// TwinCAT 3 PLC project axis_4
// ProgramVersion: 3.1.4026.27
// libraries:
//   Tc2_MC2, * (Beckhoff Automation GmbH)
//   Tc2_Standard, * (Beckhoff Automation GmbH)
//   Tc2_System, * (Beckhoff Automation GmbH)
// project tree:
//   DUTs/ ST_AxisMonitor.TcDUT, ST_MachineMonitor.TcDUT, ST_AxisCommand.TcDUT, ST_ControlStation.TcDUT, ST_AxisConfig.TcDUT, ST_TrajectoryPoint.TcDUT, ST_AxisAds.TcDUT
//   GVLs/ GVL_control.TcGVL, GVL_HMI.TcGVL, GVL_motion.TcGVL, GVL_sy.TcGVL, GVL_axis.TcGVL
//   POUs/ControlAuthority_控制权/ F_ControlDecision.TcPOU, FB_ControlAuthority.TcPOU
//   POUs/ManualControl_手动控制/ FB_AxisCommandGate.TcPOU, FB_AxisControl.TcPOU
//   POUs/Feedback_反馈/ FB_HmiFeedback.TcPOU
//   POUs/AxisConfig_轴配置/ F_AxisPositionValid.TcPOU, F_AxisConfigValid.TcPOU, FB_AxisConfig.TcPOU
//   POUs/Trajectory_点位与轨迹/ FB_FourAxisTrajectory.TcPOU, F_TrajectoryPoint.TcPOU
//   / PlcTask.TcTTO
//   POUs/ MAIN.TcPOU
// real-time tasks:
//   TASK PlcTask: cycle T#10ms, priority 20, ADS port 350
//   TASK PlcTask1: cycle T#2ms, priority 7, ADS port 351
// motion (NC):
//   TASK NC-Task 1 SAF: cycle T#2ms, priority 4, ADS port 501
//   TASK NC-Task 1 SVB: cycle T#10ms, priority 8, ADS port 511
//   AXIS axis1 (id 1)
//     OtherSettings: AllowMotionCmdToSlave=true
//     encoder EncType=19
//       EncPara: MaxCount=#xffffffff
//     drive DrvType=16
//       DrvPara: MaxCount=#xffffffff
//         Analog: TorqueSetpointScale=10, ScaleFactorActTorque=0.1
//         TimeComp: TaskDelayCycles=1
//     controller CtrType=1
//       CtrPara: PriorControlFactor=1
//         Observer: BandWidth=20
//   AXIS axis2 (id 2)
//     OtherSettings: AllowMotionCmdToSlave=true
//     encoder EncType=19
//       EncPara: MaxCount=#xffffffff
//     drive DrvType=16
//       DrvPara: MaxCount=#xffffffff
//         Analog: TorqueSetpointScale=10, ScaleFactorActTorque=0.1
//         TimeComp: TaskDelayCycles=1
//     controller CtrType=1
//       CtrPara: PriorControlFactor=1
//         Observer: BandWidth=20
//   AXIS axis3 (id 3)
//     OtherSettings: AllowMotionCmdToSlave=true
//     encoder EncType=19
//       EncPara: MaxCount=#xffffffff
//     drive DrvType=16
//       DrvPara: MaxCount=#xffffffff
//         Analog: TorqueSetpointScale=10, ScaleFactorActTorque=0.1
//         TimeComp: TaskDelayCycles=1
//     controller CtrType=1
//       CtrPara: PriorControlFactor=1
//         Observer: BandWidth=20
//   AXIS axis4 (id 4)
//     OtherSettings: AllowMotionCmdToSlave=true
//     encoder EncType=19
//       EncPara: MaxCount=#xffffffff
//     drive DrvType=16
//       DrvPara: MaxCount=#xffffffff
//         Analog: TorqueSetpointScale=10, ScaleFactorActTorque=0.1
//         TimeComp: TaskDelayCycles=1
//     controller CtrType=1
//       CtrPara: PriorControlFactor=1
//         Observer: BandWidth=20
// variable links:
//   axis_4/axis_4 Instance <-> NC-Task 1 SAF/Axes/axis1
//     PlcTask Inputs/GVL_sy.axis[1].NcToPlc <-> 输出/ToPlc
//     PlcTask Outputs/GVL_sy.axis[1].PlcToNc <-> 输入/FromPlc
//   axis_4/axis_4 Instance <-> NC-Task 1 SAF/Axes/axis2
//     PlcTask Inputs/GVL_sy.axis[2].NcToPlc <-> 输出/ToPlc
//     PlcTask Outputs/GVL_sy.axis[2].PlcToNc <-> 输入/FromPlc
//   axis_4/axis_4 Instance <-> NC-Task 1 SAF/Axes/axis3
//     PlcTask Inputs/GVL_sy.axis[3].NcToPlc <-> 输出/ToPlc
//     PlcTask Outputs/GVL_sy.axis[3].PlcToNc <-> 输入/FromPlc
//   axis_4/axis_4 Instance <-> NC-Task 1 SAF/Axes/axis4
//     PlcTask Inputs/GVL_sy.axis[4].NcToPlc <-> 输出/ToPlc
//     PlcTask Outputs/GVL_sy.axis[4].PlcToNc <-> 输入/FromPlc

CONFIGURATION axis_4
    RESOURCE PLC ON TwinCAT3
        TASK PlcTask(INTERVAL := T#2ms, PRIORITY := 7);
        PROGRAM MAIN WITH PlcTask : MAIN;
    END_RESOURCE
END_CONFIGURATION

// ---- DUTs/ST_AxisMonitor.TcDUT
{attribute 'pack_mode' := '1'}
TYPE ST_AxisMonitor :
STRUCT
    // 仅反馈，固定 22 字节；顺序与 C# PlcAxisMonitor 完全一致。
    lrActualPosition : LREAL; // PLC 从基础轴转发、上位机只读：NC 实际位置，单位跟随 NC，现场单位尚未确认。
    lrSpeed : LREAL; // PLC 从基础轴转发、上位机只读：NC 实际速度，单位为 NC 位置单位/秒，含方向正负号。
    xHomed : BOOL; // PLC 从基础轴转发、上位机只读：NC 已回原反馈，不是回原请求。
    xError : BOOL; // PLC 从基础轴转发、上位机只读：本轴 NC 或基础 MC 功能块错误。
    xPositiveLimit : BOOL; // PLC 从基础轴转发、上位机只读：正向硬限位或 NC 正向软限位超限。
    xNegativeLimit : BOOL; // PLC 从基础轴转发、上位机只读：负向硬限位或 NC 负向软限位超限。
    xOriginSignal : BOOL; // PLC 从基础轴转发、上位机只读：原点传感器信号，不代表回原已经完成。
    xEnabled : BOOL; // MC_Power.Status，使能反馈，不以运动位代替。 PLC 从基础轴转发，上位机只读。
END_STRUCT
END_TYPE

// ---- DUTs/ST_MachineMonitor.TcDUT
{attribute 'pack_mode' := '1'}
TYPE ST_MachineMonitor :
STRUCT
    // 布局版本 4，总长 164 字节；修改字段时须同步上位机并升级版本。
    nVersion : UINT; // PLC 写、上位机只读：监控协议布局版本，当前为 4，上位机据此校验帧。
    nByteSize : UINT; // PLC 写、上位机只读：完整监控结构字节数，当前为 164，不是轴数量或有效点数。
    nControlOwner : UINT; // PLC 写、上位机只读：仲裁持有者，0 未分配、1 造波控制室、2 拖车本地、3 远程操作室。
    nControlMode : UINT; // PLC 写、上位机只读：0 未分配、1 手动、2 轨迹占用；由持有者和轨迹 Busy 推导，不是模式请求。
    nWaveState : UINT; // PLC 写、上位机只读：页面状态 0 待机、1 准备、2 运行、4 停止中、5 已停止、6 完成、7 故障。
    uiWaveFaultCode : UINT; // PLC 写、上位机只读：组或首个轴的 16 位显示错误码，超过 65535 显示 65535；完整码见 GVL_HMI.udiDetailedFaultCode。
    udiHeartbeat : UDINT; // PLC 每约 500 ms 递增的反馈心跳，溢出回 0；上位机据变化判断反馈新鲜度，不由上位机写。
    Axis1 : ST_AxisMonitor; // PLC 写、上位机只读：NC 轴 1 的实际反馈，布局固定为 ST_AxisMonitor。
    Axis2 : ST_AxisMonitor; // PLC 写、上位机只读：NC 轴 2 的实际反馈，布局固定为 ST_AxisMonitor。
    Axis3 : ST_AxisMonitor; // PLC 写、上位机只读：NC 轴 3 的实际反馈，布局固定为 ST_AxisMonitor。
    Axis4 : ST_AxisMonitor; // PLC 写、上位机只读：NC 轴 4 的实际反馈，布局固定为 ST_AxisMonitor。
    // 轨迹及自动准备反馈，顺序对应 C#，继续 1 字节对齐。
    nTrajectoryState : UINT; // PLC 写、上位机只读：轨迹内部状态 0空闲/5拼表/10校验/15首点定位/20开外部给定/30运行/40末点保持/50减速/60关给定/70等停稳/90故障。
    nReceivedCount : UDINT; // PLC 写、上位机只读：四轴已登记接收的点数，也是下段起始偏移；不是已拼表点数。
    nLoadedCount : UDINT; // PLC 写、上位机只读：四轴均已拼入执行表的点数；不代表已校验通过或已运动完成。
    nPointCount : UDINT; // PLC 转发、上位机只读：上位机在 GVL_motion 中声明的目标总点数，不等于已接收或已拼接点数。
    nCurrentPoint : UDINT; // PLC 写、上位机只读：最近准备送给 NC 的点号，从 0 开始；不表示实际轴已到该点。
    udiReceivedSequence : UDINT; // PLC 写、上位机只读：当前接收表所属轨迹序号，清表后为 0；用于核对收段确认。
    udiAcceptedSequence : UDINT; // PLC 写、上位机只读：已校验通过并进入首点定位的轨迹序号，用于防止重复执行，不是完成序号。
    udiErrorId : UDINT; // PLC 写、上位机只读：轨迹块完整诊断码或 MC 原始 ErrorID；不汇总单轴错误，0 表示当前无组错误码。
    nUploadStation : UINT; // PLC 写、上位机只读：接收表归属站，0 无归属、1..3 对应控制站；不是上位机直接申请的授权。
    xUploadBusy : BOOL; // PLC 写、上位机只读：状态 5 正在统一拼表；不表示上位机当前正在写 ADS。
    xDataReady : BOOL; // PLC 写、上位机只读：完整位置表已拼接就绪；数值由上位机预检，不代表轴已使能或已到首点。
    xTrajectoryBusy : BOOL; // PLC 写、上位机只读：状态 10..70 占用轴控制，包含启动检查、定位、运行和退出；拼表状态 5 不占用。
    xRunning : BOOL; // PLC 写、上位机只读：仅内部状态 30 正常取点运行，首点定位和减速退出不算正常取点。
    xDone : BOOL; // PLC 写、上位机只读：轨迹自然完成且退出后保持，不以启动写入成功或末点已发送代替。
    xError : BOOL; // PLC 写、上位机只读：轨迹组故障保持位，确认退出并满足静止条件后由组复位请求清除。
    xStopped : BOOL; // PLC 写、上位机只读：人工组停止流程完成后保持，区别于自然完成 xDone 和组故障 xError。
    xMotionPermit : BOOL; // PLC 写、上位机只读：当前运行许可反馈，不等于已获控制权、轴已使能或硬件安全确认。
    xConfigValid : BOOL; // PLC 写、上位机只读：四轴设备参数的监控校验结果；不表示已使能或轨迹整表已校验。
    xAxesIdle : BOOL; // PLC 写、上位机只读：四轴有效停稳、基础块空闲且无外部给定；未使能轴也可满足空闲。
    xAxisFault : BOOL; // PLC 写、上位机只读：任一基础轴错误、NC 错误或 NC I/O 无效；不是仅指驱动器报警。
    xAxesStopped : BOOL; // 实际停车完成；MC_Stop 可以尚未释放。 PLC 汇总四轴 xStopped，上位机只读；反馈无效时不能确认停稳。
    // 配套版本及首次故障；均由 PLC 写，上位机只读。
    udiProgramVersion : UDINT; // PLC 源码发布号，2026102301；下载后才更新在线值。
    nBehaviorVersion : UINT; // 1=上位机整表预检，PLC 保留接收协议与运动联锁。
    nFaultAxis : UINT; // 首次轨迹故障轴号 1..4，0 表示组条件或未定位到单轴。
    nFaultSource : UINT; // 首次故障来源，含联停条件和 MC 块，见故障说明。
    nFaultState : UINT; // 首次故障发生时的轨迹阶段，不随停车阶段变化。
    udiCleanupErrorId : UDINT; // 停车/关闭/退出的首个错误，不能覆盖原始轨迹故障。
END_STRUCT
END_TYPE

// ---- DUTs/ST_AxisCommand.TcDUT
TYPE ST_AxisCommand :
STRUCT
    // 单个站点的命令邮箱，不含反馈；本站上位机写请求，PLC 在控制权交接时清空旧命令。
    xStart : BOOL; // 本站上位机写：保持型使能请求，TRUE 请求使能、FALSE 请求撤使能；不是轨迹启动或实际使能反馈。
    xStop : BOOL; // 本站上位机写：保持型停止请求，TRUE 停车、FALSE 撤请求；当前客户端发送 50 ms 脉冲，停稳另读反馈。
    jogz : BOOL; // 本站上位机写：正向点动保持位，按下 TRUE、松开 FALSE；不是实际正转反馈。
    jogf : BOOL; // 本站上位机写：负向点动保持位，按下 TRUE、松开 FALSE；不是实际反转反馈。
    gohome : BOOL; // 本站上位机写：回原上升沿请求，须先回 FALSE 再次置 TRUE；当前客户端脉冲 50 ms。
    reset : BOOL; // 本站上位机写：轴故障复位上升沿请求，须先回 FALSE 再次置 TRUE；当前客户端脉冲 50 ms。
    lrJogSpeed : LREAL; // 本站上位机写：点动速度幅值，单位为 NC 位置单位/秒；启动点动前先写速度，再写方向位。
END_STRUCT
END_TYPE

// ---- DUTs/ST_ControlStation.TcDUT
TYPE ST_ControlStation :
STRUCT
    // 站点写：先写 nAction，再提交新的非零序号；心跳独立持续更新。
    udiHeartbeat : UDINT; // 本站上位机持续写变化计数，不是请求沿；PLC 见过变化后判在线，连续 3 秒不变判离线。
    nAction : UINT; // 1 申请，2 释放。 本站上位机先写动作，再更新请求序号；动作值本身不代表已获授权。
    udiRequestSequence : UDINT; // 本站上位机写：新的非零序号提交一次请求，PLC 按与应答序号不同识别新请求，不按 BOOL 上升沿。
    xWaveSession : BOOL; // 本站发送/自动准备/执行会话，锁住交接；失联后不再保留锁。 本站写保持位，PLC 在交接时清零；表示软件会话占用，不是实际轨迹运行反馈。
    aAxis : ARRAY[1..4] OF ST_AxisCommand; // 本站上位机写：固定对应轴 1..4 的手动命令；PLC 仅转交授权站，交接时清除各站旧命令。
    // PLC 写，站点只读：请求是否成功必须看同序号应答，不能以写成功代替授权。
    udiAckSequence : UDINT; // PLC 写、本站只读：已处理的请求序号，必须等于本次请求序号后才能采用 nResult。
    nResult : UINT; // 1 成功；2 运行锁定；3 保留（旧版现场授权拒绝）；4 离线；5 非持有者；6 优先级；7 无效操作。 PLC 写、本站只读；须结合本次相同序号的 udiAckSequence 判断。
    xOnline : BOOL; // PLC 写、本站只读：心跳变化及 3 秒超时判断结果；ADS 连接成功不等于本站在线。
    xGranted : BOOL; // PLC 写、本站只读：当前持有者且在线、未失联退出时为 TRUE；写请求成功不代表获授权。
END_STRUCT
END_TYPE

// ---- DUTs/ST_AxisConfig.TcDUT
TYPE ST_AxisConfig :
STRUCT
    // 单位跟随 NC：位置、位置/秒、位置/秒²。必须按设备行程填写。
    // 参数在 FB_AxisConfig 中集中填写到 GVL_motion.aConfig；当前值仅用于虚拟轴调试，现场位置单位尚未确认。
    lrMinPosition : LREAL; // 设备配置值，PLC 读取：最小允许位置边界，单位跟随 NC 位置单位。
    lrMaxPosition : LREAL; // 设备配置值，PLC 读取：最大允许位置边界，单位跟随 NC 位置单位，须大于最小位置。
    lrMaxVelocity : LREAL; // 设备配置值，PLC 读取：点动及轨迹的速度上限，正值，单位为 NC 位置单位/秒。
    lrMaxAcceleration : LREAL; // 设备配置值，PLC 读取：点动/定位加速度及轨迹加速度幅值上限，正值，单位为 NC 位置单位/秒²。
    lrStopDeceleration : LREAL; // 设备配置值，PLC 读取：手动、首点定位及轨迹停车减速度幅值，正值且不大于最大加速度，单位为 NC 位置单位/秒²。
    lrStartTolerance : LREAL; // 设备配置值，PLC 读取：首点定位完成后实际位置和设定位置到首点的容差，轨迹要求大于 0，单位跟随 NC。
    lrInitVelocity : LREAL; // 轨迹启动前，四轴各自移动到首点的速度。 配置方填写、PLC 读取；须大于 0 且不超过最大速度，单位为 NC 位置单位/秒。
END_STRUCT
END_TYPE

// ---- DUTs/ST_TrajectoryPoint.TcDUT
TYPE ST_TrajectoryPoint :
STRUCT
    // PLC 内部送点使用；上位机只下发 LREAL 位置表，速度/加速度由相邻点计算。
    lrPosition : LREAL; // PLC 内部绝对位置给定，来自当前表点或停车积分；不是实际位置反馈，单位跟随 NC。
    lrVelocity : LREAL; // PLC 内部速度给定，正常运行由相邻点按 2 ms 中心差分计算，首尾为 0；单位为 NC 位置单位/秒。
    lrAcceleration : LREAL; // PLC 内部加速度给定，正常运行由相邻点按 2 ms 二阶差分计算，停车时另算；单位为 NC 位置单位/秒²。
END_STRUCT
END_TYPE

// ---- DUTs/ST_AxisAds.TcDUT
TYPE ST_AxisAds :
STRUCT
    // PLC → 上位机：反馈量
    lrActualPosition : LREAL; // PLC 写、上位机只读：NC 实际位置，单位跟随 NC 位置单位，现场尚未确认。
    lrSpeed          : LREAL; // PLC 写、上位机只读：NC 实际速度，单位为 NC 位置单位/秒，正负号表示方向。
    xMotorRun        : BOOL; // PLC 写、上位机只读：NC Moving 实际运动位，不是使能成功或运动请求。
    xHomed           : BOOL; // PLC 写、上位机只读：NC Homed 回原有效反馈，不以 gohome 请求代替。
    xError           : BOOL; // PLC 写、上位机只读：NC 或 Power/Stop/Home/Jog/Reset 任一错误，错误码见 udiErrorId。
    xPositiveLimit   : BOOL; // PLC 写、上位机只读：正向硬限位或 NC 正向软限位超限，TRUE 表示触发。
    xNegativeLimit   : BOOL; // PLC 写、上位机只读：负向硬限位或 NC 负向软限位超限，TRUE 表示触发。
    xOriginSignal    : BOOL; // PLC 写、上位机只读：实际原点传感器信号，不等于已完成回原。

    // PLC 命令门转交授权站的命令；上位机应写 aStation[本站].aAxis，不直写以下字段。
    xStart     : BOOL; // PLC 命令门转交：保持型使能请求，TRUE 请求使能、FALSE 先停车再撤使能；实际结果看 xEnabled。
    xStop      : BOOL; // PLC 命令门转交：保持型停止请求，TRUE 请求停车并维持停止条件，FALSE 撤请求；完成看 xStopped。
    jogz       : BOOL; // PLC 命令门转交：正向点动保持请求，按下 TRUE、释放 FALSE 后减速；与 jogf 同时 TRUE 不点动。
    jogf       : BOOL; // PLC 命令门转交：负向点动保持请求，按下 TRUE、释放 FALSE 后减速；与 jogz 同时 TRUE 不点动。
    gohome     : BOOL; // PLC 命令门转交：回原上升沿请求，须回 FALSE 后才能再次触发；完成看 xHomed。
    reset      : BOOL; // PLC 命令门转交：轴故障复位上升沿请求，须回 FALSE 后再次触发；故障是否消除看 xError。
    lrJogSpeed : LREAL; // PLC 命令门转交：点动速度幅值，单位为 NC 位置单位/秒，须大于 0 且不超过配置上限。
    // 新字段放在末尾；上位机应按 ADS 符号访问，整结构读写须同步更新布局。
    xEnabled : BOOL; // MC_Power.Status，使能反馈；xStart 为保持型使能请求。 PLC 每扫描写，上位机只读。
    xBusy : BOOL; // PLC 写、上位机只读：轨迹占用或 Jog/Home/Stop/Reset 忙，含停止锁保持，不等于轴正在运动。
    xStopped : BOOL; // 实际停稳且回原/点动退出，允许 MC_Stop.Done 保持。 PLC 写、上位机只读；不是停止请求，也不要求停止锁已经释放。
    udiErrorId : UDINT; // PLC 写、上位机只读：按 NC/Power/Stop/Home/Jog/Reset 顺序取首个错误码，0 表示未发布错误码。
END_STRUCT
END_TYPE

// ---- GVLs/GVL_control.TcGVL
{attribute 'qualified_only'}
VAR_GLOBAL
    // 新三站协议编码：1 造波控制室，2 拖车本地，3 远程操作室；数字小优先级高。
    // 各站只写自己的请求、心跳和手动命令；应答与授权结果由 PLC 写。
    aStation : ARRAY[1..3] OF ST_ControlStation; // 三站独立邮箱；各站写自己的请求/心跳/命令，PLC 写应答与授权反馈。
    // 纯软件申请，不使用现场主控选择位；PLC 按心跳、运行锁及优先级授予控制权。
    // 以下由仲裁块写，任何上位机都不能直接写 Owner 来取得权限。
    nOwner : UINT; // PLC 发布的持有站：0 未分配，1 控制室、2 拖车本地、3 远程室；上位机只读。
    xLocked : BOOL; // 统一交接锁：运动、待执行运动命令，或 I/O 故障下轴仍使能。
    xCanRelease : BOOL; // 由 Owner 和 xLocked 推导，保留此反馈供已有上位机兼容。
    xFeedbackInvalid : BOOL; // 任一轴 NC I/O 无效；单独提示，基础轴块禁止新使能/运动。
    xCanCommand : BOOL; // PLC 发布的当前持有站命令许可；需持有站在线且未失联锁存。
    xOwnerChanged : BOOL; // 本扫描发生交接或撤权重授的标志，用于清旧命令、阻止同扫描重放。
    xStopOwner : BOOL; // 失联后撤销命令并停车，保持旧 Owner 直到停稳。
END_VAR

// ---- GVLs/GVL_HMI.TcGVL
{attribute 'qualified_only'}
VAR_GLOBAL
    // 整块只读监控接口；由 FB_HmiFeedback 在轴块执行后发布。
    stMonitor : ST_MachineMonitor; // PLC 每扫描发布的整块只读监控帧，包含四轴实际状态与组反馈。
    // 保留完整故障码及轨迹诊断；全部由 PLC 发布，上位机只读。
    udiDetailedFaultCode : UDINT; // 完整错误码，不丢失高 16 位。
    nFaultAxis : UINT; // 0 为组故障或无错误；1..4 为对应轴的首个错误。
    nTrajectoryState : UINT; // 轨迹块内部 nState，区别于上述页面状态编码。
    nCurrentPoint : UDINT; // PLC 发布的最近外部给定点号，从 0 开始，不表示机械轴实际到位。
    nLoadedCount : UDINT; // PLC 发布的四轴已拼入执行表的点数。
    nPointCount : UDINT; // PLC 发布的目标单轴总点数，不表示接收或执行进度。
    xDataReady : BOOL; // PLC 发布的整表拼接完成标志，不表示数值校验或首点定位完成。
    xTrajectoryBusy : BOOL; // PLC 发布的轨迹占轴标志，含校验、定位、执行和退出阶段。
END_VAR

// ---- GVLs/GVL_motion.TcGVL
{attribute 'qualified_only'}
// ADS 协议：上位机写命令/数据，PLC 写反馈；状态字段只供上位机读取。
// PC 连续提交各段，全部下发后用 xAssemble 请求 PLC 拼表；xDataReady 后才允许启动。
// xUpload/xAssemble/xClear/xStart/xReset 都需回 FALSE 后再产生下一次上升沿。
VAR_GLOBAL
    // 运行许可由 MAIN 每扫描写入；当前仅用于虚拟轴调试。
    xMotionPermit : BOOL; // 实机改接安全继电器允许反馈，不代替硬件安全回路。
    axPositiveLimit : ARRAY[1..4] OF BOOL; // 四轴正向硬限位输入，索引为轴号 1～4，TRUE 表示触发。
    axNegativeLimit : ARRAY[1..4] OF BOOL; // 四轴负向硬限位输入，索引为轴号 1～4，TRUE 表示触发。
    axHomeSensor : ARRAY[1..4] OF BOOL; // 四轴原点开关输入，索引为轴号 1～4，传给 NC 标准回零校准凸轮。
    // 四轴配置只在 FB_AxisConfig 中填写，手动、反馈和轨迹均读取此数组。
    aConfig : ARRAY[1..4] OF ST_AxisConfig; // 单位跟随 NC；空闲时由配置块直接更新，运动期间保持。

    // 以下为上位机写入的轨迹命令与点位；nUploadStation、xStopped 两项由 PLC 写、上位机只读。
    nCommandStation : UINT; // 上位机命令来源，必须等于有效 Owner；不是授权本身。
    nUploadStation : UINT; // PLC 锁存的上传所属站，只读。
    xStopped : BOOL; // 人工停止完成；不同于自然完成 xDone 或故障。
    // 参考旧工程的独立分段区：21 段、每段四轴、每轴最多 100000 个 LREAL 点。
    // 下标依次为 [段号, 轴号, 段内点号]；已提交段禁止覆盖，全部下发后统一拼接。
    aUpload : ARRAY[0..20, 1..4, 0..99999] OF LREAL; // 上位机写入的独立位置段：[段0～20,轴1～4,段内点0～99999]，数值单位跟随 NC。
    nPointCount : UDINT; // 整条轨迹总点数，4..2100000。
    nSampleTimeUs : UINT := 2000; // 单位微秒，目前仅接受 2000。
    udiUploadSequence : UDINT; // 整条轨迹使用同一个非零序号。
    nUploadOffset : UDINT; // 本段全局偏移，必须等于 nReceivedCount，段号=偏移/100000。
    nUploadCount : UDINT; // 非末段必须 100000 点；末段为总点数的剩余量。
    xUpload : BOOL; // 四轴本段数据写完后上升沿登记，只确认接收，不拼表。
    xAssemble : BOOL; // 全部段确认后上升沿请求统一拼表；拼接期间所有段保持不变。
    xClear : BOOL; // 空闲时上升沿清除整条位置表的就绪状态，开始新一轮上传。
    xStart : BOOL; // 完整位置表到齐后，上升沿启动。
    xStop : BOOL; // 保持型组停止，启动前必须释放。
    xReset : BOOL; // 清组故障；各轴故障用 Axis1..4.reset。
    udiHeartbeat : UDINT; // 校验/运动期间 1 秒不变化则联停。

    // 以下字段由 PLC 写，上位机只读。
    nReceivedCount : UDINT; // 已登记的下发点数，也是下一段允许的起始偏移；不代表已拼接。
    udiReceivedSequence : UDINT; // 已登记各段所属轨迹序号，清表后为 0。
    xUploadBusy : BOOL; // 全部下发后的统一拼表正在执行，不表示 PC 正在写 ADS。
    nLoadedCount : UDINT; // 四轴均已拼入完整表的点数；下发期间始终为 0。
    xDataReady : BOOL; // 全部段已统一拼接完成，不表示已校验或已定位到首点。
    xBusy : BOOL; // 校验、首点定位、执行和退出期间占用轴控制。
    xRunning : BOOL; // 状态 30，首点定位及减速不算正常取点运行。
    xDone : BOOL; // 正常完成后保持，清表/复位/新启动时清除。
    xError : BOOL; // 组故障保持位，需确认退出和静止后复位。
    udiErrorId : UDINT; // 首次故障的程序诊断码或 MC 原始 ErrorID，详见说明文档。
    nFaultAxis : UINT; // 首次故障轴 1..4；组故障或无故障为 0，复位时清除。
    nFaultSource : UINT; // 首次故障来源：1许可/2控制权/3使能/4单轴停止/5手动冲突/6限位，7..20见故障说明。
    nFaultState : UINT; // 首次故障发生阶段；故障退出期间保持，不能用当前停车阶段替代。
    udiCleanupErrorId : UDINT; // 首个停车、关闭或退出错误，保留原始 udiErrorId。
    nState : UINT; // 对应轨迹块 CASE 的 0/5/10/15/20/30/40/50/60/70/90。
    nCurrentPoint : UDINT; // 最近送出的点号，0 起始。
    udiAcceptedSequence : UDINT; // 已进入首点定位的轨迹序号，不能重复执行。
END_VAR

// ---- GVLs/GVL_sy.TcGVL
VAR_GLOBAL

axis  : ARRAY[1..4] OF AXIS_REF; // 四根 NC 轴引用，固定索引 1～4；轴状态从 NC 读取，运动块经此接口下发控制。

END_VAR

// ---- GVLs/GVL_axis.TcGVL
VAR_GLOBAL
    // PLC 内部手动命令与轴反馈；命令由 A03_ManualCommands 转交，反馈由基础轴块更新。
    // 上位机手动命令写 GVL_control.aStation[站号].aAxis，状态读取 GVL_HMI.stMonitor。

    Axis1 : ST_AxisAds; // 轴1内部手动命令与实际反馈；命令由命令门转交，反馈由轴1基础块更新。
    Axis2 : ST_AxisAds; // 轴2内部手动命令与实际反馈；命令由命令门转交，反馈由轴2基础块更新。
    Axis3 : ST_AxisAds; // 轴3内部手动命令与实际反馈；命令由命令门转交，反馈由轴3基础块更新。
    Axis4 : ST_AxisAds; // 轴4内部手动命令与实际反馈；命令由命令门转交，反馈由轴4基础块更新。


END_VAR

// ---- POUs/MAIN.TcPOU
// PlcTask 每 2 ms 调用；先刷新反馈，再判组条件，再轨迹，最后基础轴块。
// 每轴的 NC 引用、ADS 数据、参数及传感器索引必须一一对应。
PROGRAM MAIN
VAR
    fbAxisConfig : FB_AxisConfig; // 独立轴配置入口，仅在有效空闲时应用本块的虚拟轴参数。
    fbAxis1 : FB_AxisControl; // 轴1基础控制实例，固定对应 GVL_sy.axis[1] 和 GVL_axis.Axis1。
    fbAxis2 : FB_AxisControl; // 轴2基础控制实例，固定对应 GVL_sy.axis[2] 和 GVL_axis.Axis2。
    fbAxis3 : FB_AxisControl; // 轴3基础控制实例，固定对应 GVL_sy.axis[3] 和 GVL_axis.Axis3。
    fbAxis4 : FB_AxisControl; // 轴4基础控制实例，固定对应 GVL_sy.axis[4] 和 GVL_axis.Axis4。
    fbAuthority : FB_ControlAuthority; // 三站控制权仲裁实例，处理申请、释放、心跳和交接锁。
    aCommandGate : ARRAY[1..4] OF FB_AxisCommandGate; // 四轴手动命令门，只向对应轴转交当前持有站的有效命令。
    xControlBusy : BOOL; // 实际运动、轨迹或轴块忙的汇总，作为禁止控制权交接的判据。
    nManualStation : UINT; // 本扫描允许读取的站号；0 时命令门清除旧请求。
    fbTrajectory : FB_FourAxisTrajectory; // 四轴点位接收、拼表、校验及轨迹执行实例。
    fbHmiFeedback : FB_HmiFeedback; // 四轴执行结果发布到 switch 只读监控接口。
    xAllEnabled : BOOL; // 四轴使能反馈，用于运行中判断是否掉使能。
    xAxesReady : BOOL; // 轨迹启动就绪：四轴使能、回原、静止且不在停车。
    nAbortReason : UINT; // 本扫描首个联停原因；0 表示没有联停请求。
    xAbort : BOOL; // 整组联停请求，汇总许可丢失、撤使能、命令冲突及限位等条件。
    xAxisFault : BOOL; // 任一基础轴错误或 NC 错误、I/O 无效，供轨迹块判断故障。
    i : INT; // 四轴状态汇总的循环轴号，范围 1～4。
END_VAR

// 当前仅用于虚拟轴软件调试，明确给出运行许可。
// 接实机前必须将下一行替换为现场安全继电器的运行允许反馈。
GVL_motion.xMotionPermit := TRUE;

// 刷新四轴实际状态；只读取 NC 反馈，不要求持有控制权。
A01_ReadAxisStatus();

// 汇总交接条件并处理控制权；写入 GVL_control 仲裁反馈。
A02_ControlAuthority();

// 轴配置单独处理，使用当前运动锁和现有空闲反馈。
fbAxisConfig();

// 取出授权站手动命令；通过命令门写入 GVL_axis 命令字段。
A03_ManualCommands();

// 汇总轨迹联锁并调用原轨迹块；更新 GVL_motion 轨迹状态。
A04_TrajectoryControl();

// 调用四轴基础控制；更新 NC 控制输出及 GVL_axis 实际反馈。
A05_ManualAxes();

// 发布本扫描执行后的反馈；只写 GVL_HMI，不产生运动命令。
A06_PublishFeedback();

ACTION A01_ReadAxisStatus:
// 刷新四轴实际状态；只读取 NC 反馈，不要求持有控制权。
// 先统一刷新轴状态，再决定四轴本周期的共同轨迹帧。
FOR i := 1 TO 4 DO
 GVL_sy.axis[i].ReadStatus();
 END_FOR
END_ACTION

ACTION A02_ControlAuthority:
// 汇总交接条件并处理控制权；写入 GVL_control 仲裁反馈。
// 运行锁：点动、回原、轨迹、停止/退出及未消费的运动命令都阻止交接。
// 使用 NC 状态、实际速度和轴块 Busy；I/O 无效单独发布，不能冒充运动占用。
xControlBusy := GVL_motion.xBusy OR GVL_axis.Axis1.xBusy OR GVL_axis.Axis2.xBusy
    OR GVL_axis.Axis3.xBusy OR GVL_axis.Axis4.xBusy;
GVL_control.xFeedbackInvalid := FALSE;
FOR i := 1 TO 4 DO
    xControlBusy := xControlBusy OR GVL_sy.axis[i].Status.Moving
        OR GVL_sy.axis[i].Status.Homing OR GVL_sy.axis[i].Status.Stopping
        OR GVL_sy.axis[i].Status.ExtSetPointGenEnabled
        OR (ABS(GVL_sy.axis[i].NcToPlc.ActVelo) > 0.000001);
    GVL_control.xFeedbackInvalid := GVL_control.xFeedbackInvalid OR GVL_sy.axis[i].Status.IoDataInvalid;
END_FOR
fbAuthority(xMotionBusy := xControlBusy, xFeedbackInvalid := GVL_control.xFeedbackInvalid);
END_ACTION

ACTION A03_ManualCommands:
// 四个命令门共用本扫描的授权结果，各自读取对应轴的邮箱。
// 交接扫描仍清除旧请求，新持有者须在确认授权后重新发命令。
nManualStation := 0;
IF GVL_control.xCanCommand AND NOT GVL_control.xOwnerChanged THEN
    nManualStation := GVL_control.nOwner;
END_IF
aCommandGate[1](Data := GVL_axis.Axis1, nStation := nManualStation, nAxis := 1, xStop := GVL_control.xStopOwner);
aCommandGate[2](Data := GVL_axis.Axis2, nStation := nManualStation, nAxis := 2, xStop := GVL_control.xStopOwner);
aCommandGate[3](Data := GVL_axis.Axis3, nStation := nManualStation, nAxis := 3, xStop := GVL_control.xStopOwner);
aCommandGate[4](Data := GVL_axis.Axis4, nStation := nManualStation, nAxis := 4, xStop := GVL_control.xStopOwner);
END_ACTION

ACTION A04_TrajectoryControl:
// 汇总轨迹联锁并调用原轨迹块；更新 GVL_motion 轨迹状态。
// 基础轴块在轨迹块之后调用，此处使用上一扫描的使能反馈。
xAllEnabled := GVL_axis.Axis1.xEnabled AND GVL_axis.Axis2.xEnabled AND GVL_axis.Axis3.xEnabled AND GVL_axis.Axis4.xEnabled;
xAxisFault := GVL_axis.Axis1.xError OR GVL_axis.Axis2.xError  OR GVL_axis.Axis3.xError OR GVL_axis.Axis4.xError;
// 按许可、控制权、使能、停止、手动冲突、限位的顺序取第一个联停原因。
// 当前持有站发出的整组停止命令，由轨迹块走正常停车流程。
nAbortReason := 0;
IF NOT GVL_motion.xMotionPermit THEN nAbortReason := 1;
ELSIF NOT GVL_control.xCanCommand THEN nAbortReason := 2;
ELSIF (GVL_motion.xBusy AND NOT xAllEnabled)
    OR NOT GVL_axis.Axis1.xStart OR NOT GVL_axis.Axis2.xStart
    OR NOT GVL_axis.Axis3.xStart OR NOT GVL_axis.Axis4.xStart THEN nAbortReason := 3;
ELSIF (GVL_axis.Axis1.xStop OR GVL_axis.Axis2.xStop OR GVL_axis.Axis3.xStop OR GVL_axis.Axis4.xStop)
    AND NOT ((GVL_motion.nCommandStation = GVL_control.nOwner) AND GVL_motion.xStop) THEN nAbortReason := 4;
ELSIF GVL_axis.Axis1.jogz OR GVL_axis.Axis1.jogf OR GVL_axis.Axis1.gohome OR GVL_axis.Axis1.reset
    OR GVL_axis.Axis2.jogz OR GVL_axis.Axis2.jogf OR GVL_axis.Axis2.gohome OR GVL_axis.Axis2.reset
    OR GVL_axis.Axis3.jogz OR GVL_axis.Axis3.jogf OR GVL_axis.Axis3.gohome OR GVL_axis.Axis3.reset
    OR GVL_axis.Axis4.jogz OR GVL_axis.Axis4.jogf OR GVL_axis.Axis4.gohome OR GVL_axis.Axis4.reset THEN
    nAbortReason := 5;
END_IF
// 启动就绪才要求回原和静止，运行中用使能反馈判断掉使能。
xAxesReady := xAllEnabled;
FOR i := 1 TO 4 DO
    xAxesReady := xAxesReady AND GVL_sy.axis[i].Status.Homed AND GVL_sy.axis[i].Status.StandStill AND NOT GVL_sy.axis[i].Status.Stopping;
    xAxisFault := xAxisFault OR GVL_sy.axis[i].Status.Error OR GVL_sy.axis[i].Status.IoDataInvalid;
    IF (nAbortReason = 0) AND (GVL_motion.axPositiveLimit[i] OR GVL_motion.axNegativeLimit[i]
        OR GVL_sy.axis[i].Status.SoftLimitMinExceeded OR GVL_sy.axis[i].Status.SoftLimitMaxExceeded) THEN
        nAbortReason := 6;
    END_IF
END_FOR
xAbort := nAbortReason <> 0;
// 轨迹块先更新组状态和 xBusy，后面的基础块在本扫描就能据此禁止手动抢占。
// 全部下发后的统一拼表状态 5 不置 xBusy，不占用基础轴控制。
fbTrajectory(Axes := GVL_sy.axis, xAxesReady := xAxesReady, xAbort := xAbort, xAxisFault := xAxisFault, nAbortReason := nAbortReason);
END_ACTION

ACTION A05_ManualAxes:
// 调用四轴基础控制；更新 NC 控制输出及 GVL_axis 实际反馈。
// 四个实例各自保存 Power/Jog/Home/Stop/Reset 的状态，便于逐轴打断点。
// 四个基础实例每扫描都调用，持续更新异步 MC 块 Busy/Done/Error。
// Axis1..4 固定对应 NC 引用 [1]..[4]，不通过选中轴号复用一个实例。
fbAxis1(Axis := GVL_sy.axis[1], Data := GVL_axis.Axis1, Config := GVL_motion.aConfig[1],
    xPermit := GVL_motion.xMotionPermit AND GVL_control.xCanCommand, xPositiveLimit := GVL_motion.axPositiveLimit[1],
    xNegativeLimit := GVL_motion.axNegativeLimit[1], xHomeSensor := GVL_motion.axHomeSensor[1],
    xGroupBusy := GVL_motion.xBusy);
fbAxis2(Axis := GVL_sy.axis[2], Data := GVL_axis.Axis2, Config := GVL_motion.aConfig[2],
    xPermit := GVL_motion.xMotionPermit AND GVL_control.xCanCommand, xPositiveLimit := GVL_motion.axPositiveLimit[2],
    xNegativeLimit := GVL_motion.axNegativeLimit[2], xHomeSensor := GVL_motion.axHomeSensor[2],
    xGroupBusy := GVL_motion.xBusy);
fbAxis3(Axis := GVL_sy.axis[3], Data := GVL_axis.Axis3, Config := GVL_motion.aConfig[3],
    xPermit := GVL_motion.xMotionPermit AND GVL_control.xCanCommand, xPositiveLimit := GVL_motion.axPositiveLimit[3],
    xNegativeLimit := GVL_motion.axNegativeLimit[3], xHomeSensor := GVL_motion.axHomeSensor[3],
    xGroupBusy := GVL_motion.xBusy);
fbAxis4(Axis := GVL_sy.axis[4], Data := GVL_axis.Axis4, Config := GVL_motion.aConfig[4],
    xPermit := GVL_motion.xMotionPermit AND GVL_control.xCanCommand, xPositiveLimit := GVL_motion.axPositiveLimit[4],
    xNegativeLimit := GVL_motion.axNegativeLimit[4], xHomeSensor := GVL_motion.axHomeSensor[4],
    xGroupBusy := GVL_motion.xBusy);
END_ACTION

ACTION A06_PublishFeedback:
// 发布本扫描执行后的反馈；只写 GVL_HMI，不产生运动命令。
// 所有基础块本周期输出更新后，再发布 HMI 状态；避免把请求位误当成执行反馈。
fbHmiFeedback();
END_ACTION

END_PROGRAM

// ---- POUs/AxisConfig_轴配置/FB_AxisConfig.TcPOU
FUNCTION_BLOCK FB_AxisConfig
// 轴配置单独在此填写，直接写入全局四轴参数。
// 当前值仅用于虚拟轴调试；接实机时须按实际 NC 单位、行程和动态参数重新配置。
VAR
    i : INT; // 四轴配置下标，1～4；复用已有状态反馈，不另存初始化或空闲标志。
END_VAR

// 空闲反馈来自上一扫描；当前扫描的运动锁和 I/O 有效性由 MAIN 的 A02 更新。
// 等待有效停稳、轴块/轨迹/拼表空闲，以及点动、回原、轨迹启动请求释放。
IF GVL_HMI.stMonitor.xAxesIdle AND NOT GVL_control.xLocked AND NOT GVL_control.xFeedbackInvalid
    AND NOT GVL_motion.xBusy AND NOT GVL_motion.xUploadBusy AND NOT GVL_motion.xStart
    // 再直接确认当前 NC 停稳，避免使用上扫描空闲值时漏掉新出现的无效速度。
    AND (GVL_sy.axis[1].Status.StandStill OR GVL_sy.axis[1].Status.Disabled)
    AND (GVL_sy.axis[2].Status.StandStill OR GVL_sy.axis[2].Status.Disabled)
    AND (GVL_sy.axis[3].Status.StandStill OR GVL_sy.axis[3].Status.Disabled)
    AND (GVL_sy.axis[4].Status.StandStill OR GVL_sy.axis[4].Status.Disabled)
    AND (ABS(GVL_sy.axis[1].NcToPlc.ActVelo) <= 0.000001)
    AND (ABS(GVL_sy.axis[2].NcToPlc.ActVelo) <= 0.000001)
    AND (ABS(GVL_sy.axis[3].NcToPlc.ActVelo) <= 0.000001)
    AND (ABS(GVL_sy.axis[4].NcToPlc.ActVelo) <= 0.000001) THEN
    FOR i := 1 TO 4 DO
        // 当前四根虚拟轴使用相同参数，空闲时直接应用本块数值，已有旧值也能更新。
        // 200/12000 按本次虚拟轴调试确认；不作为实机速度、加速度能力。
        GVL_motion.aConfig[i].lrMinPosition := -200;
        GVL_motion.aConfig[i].lrMaxPosition := 200;
        GVL_motion.aConfig[i].lrMaxVelocity := 200;
        GVL_motion.aConfig[i].lrMaxAcceleration := 12000;
        GVL_motion.aConfig[i].lrStopDeceleration := 100;
        GVL_motion.aConfig[i].lrInitVelocity := 10;
        GVL_motion.aConfig[i].lrStartTolerance := 10;
    END_FOR
END_IF

END_FUNCTION_BLOCK

// ---- POUs/ManualControl_手动控制/FB_AxisControl.TcPOU
FUNCTION_BLOCK FB_AxisControl
// 单轴基础控制：使能、复位、手动点动、标准回原、停止及反馈。
// 四轴分别使用独立实例；本块不读取位置表，轨迹块通过 xGroupBusy 占用轴控制。
VAR_INPUT
    xPermit : BOOL; // 普通运行及控制权许可；FALSE 请求停车，并禁止新使能和新手动动作。
    xPositiveLimit : BOOL; // 正向硬限位，TRUE 表示触发。
    xNegativeLimit : BOOL; // 负向硬限位，TRUE 表示触发。
    xHomeSensor : BOOL; // 实际原点开关，作为标准回原校准凸轮信号。
    xGroupBusy : BOOL; // 轨迹占用时禁止手动点动、回原和复位抢占。
    Config : ST_AxisConfig; // 本轴行程及动态参数，单位跟随 NC。
END_VAR
VAR_IN_OUT
    Axis : AXIS_REF; // 对应 NC 轴引用，直接操作原轴接口。
    Data : ST_AxisAds; // 内部轴命令及反馈；命令由命令门转交，本块读取命令并更新实际反馈。
END_VAR
VAR
    fbPower : MC_Power; // 轴软件使能实例；Status 才是实际使能反馈，Data.xStart 仅为请求。
    fbJog : MC_Jog; // 正反点动实例；速度单位为 NC 位置单位/秒。
    fbHome : MC_Home; // NC 标准回零实例，使用配置的回零方式和原点凸轮信号。
    fbStop : MC_Stop; // 单轴减速停止实例；Execute 释放后仍需等待 Busy 解锁。
    fbReset : MC_Reset; // NC 轴报警复位实例，不代替运动块或轨迹组的独立故障复位。
    rtHome : R_TRIG; // 回零请求上升沿检测，输入保持 TRUE 不重复发起回零。
    rtReset : R_TRIG; // 轴复位请求上升沿检测，输入保持 TRUE 不重复发起复位。
    xPositionValid : BOOL; // 位置范围单独校验，只用于方向限制。
    xConfigValid : BOOL; // 运动参数校验，只限制点动/回原，不限制基础使能。
    xManual : BOOL; // 允许手动运动的公共条件。
    xStopRequest : BOOL; // 停止、撤使能、许可丢失、限位或运动中参数失效产生的停车条件。
    xHoldPower : BOOL; // 运动/停车未完成或组仍占用时，临时保持已有使能。
    xJogArmed : BOOL; // 联停或轨迹占用后，须先释放按钮才重新允许点动。
    xJogSpeedValid : BOOL; // 点动速度为正且不超过最大速度。
    lrJogVelocity : LREAL; // 本扫描合法点动速度，单位为 NC 位置单位/秒；无效输入置零。
    lrStopDeceleration : LREAL; // 本扫描停车减速度，单位为 NC 位置单位/秒²；参数无效时按 MC_Stop 默认规则处理。
END_VAR

// ReadStatus 在 MAIN 开头统一执行，所有轴使用本周期反馈。
// 1. 回原/复位取上升沿；输入保持 TRUE 不会每扫描重复发起。
rtHome(CLK := Data.gohome);
rtReset(CLK := Data.reset);
// Config 由 MAIN 传入 GVL_motion.aConfig；本块只读取，不覆盖输入参数。
// 2. 分开校验位置和运动参数；未配置时可以基础使能，但不允许发起运动。
xPositionValid := F_AxisPositionValid(Config);
xConfigValid := F_AxisConfigValid(Config);

// 3. 软件使能：Data.xStart 是持续使能请求，xPermit 和有效 I/O 决定能否接受该请求。
// 已经使能的轴在运动、轨迹占用或 MC_Stop 尚未结束时，由 xHoldPower 暂时保持使能。
// MC_Power 先执行，下面的 MC_Stop 使用本扫描更新后的使能反馈。
xHoldPower := fbPower.Status AND (Axis.Status.Moving OR xGroupBusy
    OR (fbStop.Busy AND NOT fbStop.Done AND NOT fbStop.Error));
// 正负方向受硬限位约束，位置范围有效时再检查位置边界。
fbPower(Axis := Axis, Enable := (Data.xStart AND xPermit AND NOT Axis.Status.IoDataInvalid) OR xHoldPower,
    Enable_Positive := NOT xPositiveLimit AND (NOT xPositionValid OR (Axis.NcToPlc.ActPos < Config.lrMaxPosition)),
    Enable_Negative := NOT xNegativeLimit AND (NOT xPositionValid OR (Axis.NcToPlc.ActPos > Config.lrMinPosition)), Override := 100);

// 4. 停车请求：停止、撤使能、许可丢失、限位或运动中参数失效。
xStopRequest := Data.xStop OR NOT Data.xStart OR NOT xPermit OR xPositiveLimit OR xNegativeLimit
    OR (NOT xConfigValid AND (Axis.Status.Moving OR fbJog.Busy OR fbHome.Busy));
// 配置无效也必须能停车；0 按 MC_Stop 默认规则沿用最近运动命令的减速度。
lrStopDeceleration := 0;
IF xConfigValid THEN lrStopDeceleration := Config.lrStopDeceleration; END_IF
// 轨迹占用或外部给定仍开启时，由轨迹块负责停车。
// MC_Stop 的 Execute 释放后，等 Busy 变为 FALSE 才允许新的手动运动。
fbStop(Axis := Axis, Execute := xStopRequest AND fbPower.Status
    AND NOT xGroupBusy AND NOT Axis.Status.ExtSetPointGenEnabled,
    Deceleration := lrStopDeceleration);

// 5. 新手动动作许可：本扫描的使能、停车和反馈状态共同决定能否点动或回原。
// Data.reset 同时阻断手动，避免同一扫描复位和点动并发。
xManual := xPermit AND xConfigValid AND fbPower.Status AND NOT xStopRequest
    AND NOT xGroupBusy AND NOT Axis.Status.ExtSetPointGenEnabled
    AND NOT fbStop.Busy AND NOT Axis.Status.Error AND NOT Axis.Status.IoDataInvalid
    AND NOT fbReset.Busy AND NOT Data.reset;
// 6. 上位机主动复位；本块不自动反复复位故障轴。
fbReset(Axis := Axis, Execute := rtReset.Q AND NOT xGroupBusy
    AND NOT Axis.Status.Moving AND NOT Data.xStop);
// 7. MC_DefaultHoming 使用 NC 配置的回原方式、速度和参考位置。
// 原点输入接实际传感器；点动按钮释放且点动块不忙时才允许启动回原。
fbHome(Axis := Axis, Execute := rtHome.Q AND xManual
    AND NOT fbJog.Busy AND NOT Data.jogz AND NOT Data.jogf,
    HomingMode := MC_DefaultHoming, bCalibrationCam := xHomeSensor);
// 正反同时按下不点动；释放按钮由 MC_Jog 按 NC 参数减速。
// 联停或轨迹占用后，必须先释放点动按钮，防止旧命令自动恢复运动。
IF NOT xManual OR fbHome.Busy THEN xJogArmed := FALSE;
ELSIF NOT Data.jogz AND NOT Data.jogf THEN xJogArmed := TRUE;
END_IF
xJogSpeedValid := (Data.lrJogSpeed > 0) AND (Data.lrJogSpeed <= Config.lrMaxVelocity);
lrJogVelocity := 0;
IF xJogSpeedValid THEN lrJogVelocity := Data.lrJogSpeed; END_IF
// 8. jogz 正向、jogf 负向，保持运行、释放减速；正反同时按下不运行。
// CONTINOUS 是 Tc2_MC2 的实际枚举名称，采用这里传入的速度和动态参数。
fbJog(Axis := Axis, JogForward := Data.jogz AND NOT Data.jogf
    AND xManual AND xJogArmed AND xJogSpeedValid AND NOT fbHome.Busy AND NOT Data.gohome,
    JogBackwards := Data.jogf AND NOT Data.jogz
    AND xManual AND xJogArmed AND xJogSpeedValid AND NOT fbHome.Busy AND NOT Data.gohome,
    Mode := MC_JOGMODE_CONTINOUS, // Tc2_MC2 的枚举名称使用 CONTINOUS 拼写。
    Velocity := lrJogVelocity,
    Acceleration := Config.lrMaxAcceleration, Deceleration := Config.lrStopDeceleration);

// 9. 反馈来源为 NC 实际状态和 MC 输出，不用上位机请求位代替执行结果。
// xEnabled=Power.Status，xHomed=NC.Homed；ErrorID 依 NC/Power/Stop/Home/Jog/Reset 顺序取首项。
Data.lrActualPosition := Axis.NcToPlc.ActPos;
Data.lrSpeed := Axis.NcToPlc.ActVelo;
Data.xMotorRun := Axis.Status.Moving;
Data.xEnabled := fbPower.Status;
Data.xHomed := Axis.Status.Homed;
Data.xPositiveLimit := xPositiveLimit OR Axis.Status.SoftLimitMaxExceeded;
Data.xNegativeLimit := xNegativeLimit OR Axis.Status.SoftLimitMinExceeded;
Data.xOriginSignal := xHomeSensor;
// MC_Stop Execute 保持时 Busy 可持续为 TRUE；停车确认与块释放分开反馈。
Data.xStopped := NOT Axis.Status.Moving AND NOT Axis.Status.IoDataInvalid
    AND (ABS(Axis.NcToPlc.ActVelo) <= 0.000001) AND NOT fbJog.Busy AND NOT fbHome.Busy
    AND NOT fbReset.Busy AND (NOT fbStop.Busy OR fbStop.Done);
Data.xBusy := xGroupBusy OR fbJog.Busy OR fbHome.Busy OR fbStop.Busy OR fbReset.Busy;
Data.udiErrorId := 0;
IF Axis.Status.Error THEN Data.udiErrorId := Axis.Status.ErrorId;
ELSIF fbPower.Error THEN Data.udiErrorId := fbPower.ErrorID;
ELSIF fbStop.Error THEN Data.udiErrorId := fbStop.ErrorID;
ELSIF fbHome.Error THEN Data.udiErrorId := fbHome.ErrorID;
ELSIF fbJog.Error THEN Data.udiErrorId := fbJog.ErrorID;
ELSIF fbReset.Error THEN Data.udiErrorId := fbReset.ErrorID;
END_IF
Data.xError := Axis.Status.Error OR fbPower.Error OR fbStop.Error
    OR fbHome.Error OR fbJog.Error OR fbReset.Error;

END_FUNCTION_BLOCK

// ---- POUs/AxisConfig_轴配置/F_AxisPositionValid.TcPOU
FUNCTION F_AxisPositionValid : BOOL
VAR_INPUT
    Config : ST_AxisConfig; // 本轴参数，只读取调用方传入的值。
END_VAR

// 只校验位置范围，供手动方向限制使用。
F_AxisPositionValid := (Config.lrMinPosition >= -1.0E12) AND (Config.lrMaxPosition <= 1.0E12)
    AND (Config.lrMinPosition < Config.lrMaxPosition);

END_FUNCTION

// ---- POUs/AxisConfig_轴配置/F_AxisConfigValid.TcPOU
FUNCTION F_AxisConfigValid : BOOL
VAR_INPUT
    Config : ST_AxisConfig; // 本轴参数，只读取调用方传入的值。
END_VAR

// 基础运动参数共用规则；首点速度和到位容差由调用方按用途检查。
F_AxisConfigValid := F_AxisPositionValid(Config)
    AND (Config.lrMaxVelocity > 0) AND (Config.lrMaxVelocity < 1.0E12)
    AND (Config.lrMaxAcceleration > 0) AND (Config.lrMaxAcceleration < 1.0E12)
    AND (Config.lrStopDeceleration > 0)
    AND (Config.lrStopDeceleration <= Config.lrMaxAcceleration);

END_FUNCTION

// ---- POUs/ControlAuthority_控制权/FB_ControlAuthority.TcPOU
FUNCTION_BLOCK FB_ControlAuthority
VAR_INPUT
    xMotionBusy : BOOL; // 含实际运动、轨迹占用、轴块 Busy，不仅看造波运行位。
    xFeedbackInvalid : BOOL; // I/O 故障只在轴仍使能时阻止交接，未使能时可申请和释放。
END_VAR
VAR
    nOwner : UINT; // 私有持有者，启动 0；GVL_control.nOwner 只是只读发布副本。
    nOldOwner : UINT; // 本扫描开始时的持有站，用于识别本扫描是否发生控制权交接。
    xOwnerLost : BOOL; // 持有站失联锁存；恢复心跳不恢复旧授权，停稳后才清旧持有者。
    xResetCommands : BOOL; // 撤权后同扫描重新授予原站，也必须清旧命令。
    xLocked : BOOL; // 申请、释放、失联退出统一使用这一份运动联锁。
    axSeenHeartbeat : ARRAY[1..3] OF BOOL; // 各站自启动以来是否出现过心跳变化，索引 1～3 对应站号。
    aLastHeartbeat : ARRAY[1..3] OF UDINT; // 各站上一扫描心跳值，仅用于判断心跳是否变化，不要求连续递增。
    aTimeout : ARRAY[1..3] OF TON; // 各站心跳超时定时器；连续 3 秒不变化判离线。
    aEmpty : ARRAY[1..4] OF ST_AxisCommand; // 四轴全零命令模板，交接时清各站旧命令，防止动作重放。
    i : INT; // 站点循环索引，范围 1～3。
    j : INT; // 当前站手动命令的轴索引，范围 1～4。
    nReply : UINT; // 本次仲裁应答码：1 成功、2 锁定、4 离线、5 非持有者、6 优先级、7 无效请求。
END_VAR

nOldOwner := nOwner;
xResetCommands := FALSE;
FOR i := 1 TO 3 DO
    IF GVL_control.aStation[i].udiHeartbeat <> aLastHeartbeat[i] THEN axSeenHeartbeat[i] := TRUE; END_IF
    aTimeout[i](IN := GVL_control.aStation[i].udiHeartbeat = aLastHeartbeat[i], PT := T#3S);
    aLastHeartbeat[i] := GVL_control.aStation[i].udiHeartbeat;
    GVL_control.aStation[i].xOnline := axSeenHeartbeat[i] AND NOT aTimeout[i].Q;
END_FOR
// 纯软件申请：三站均可申请，由在线状态、运行锁和站号优先级决定结果。

// 一份联锁：有运动占用，或 I/O 故障且轴仍使能时，禁止交接。
// I/O 故障本身不锁控制权；基础轴块仍独立禁止故障下的新使能和运动。
xLocked := xMotionBusy OR (xFeedbackInvalid AND (GVL_axis.Axis1.xEnabled
    OR GVL_axis.Axis2.xEnabled OR GVL_axis.Axis3.xEnabled OR GVL_axis.Axis4.xEnabled));
IF nOwner <> 0 THEN
    IF NOT GVL_control.aStation[nOwner].xOnline THEN xOwnerLost := TRUE; END_IF
    // 已接收但尚未进入 NC 运动的命令也锁住交接，覆盖“申请与启动同一扫描”的窗口。
    // 失联后忽略旧邮箱中的保持命令，让实际停车完成后可以退出，不会永远卡住 Owner。
    IF NOT xOwnerLost THEN
        FOR j := 1 TO 4 DO
            xLocked := xLocked OR GVL_control.aStation[nOwner].aAxis[j].jogz
                OR GVL_control.aStation[nOwner].aAxis[j].jogf
                OR GVL_control.aStation[nOwner].aAxis[j].gohome;
        END_FOR
        xLocked := xLocked OR GVL_control.aStation[nOwner].xWaveSession
            OR ((GVL_motion.nCommandStation = nOwner) AND GVL_motion.xStart);
    END_IF
    // 失联先撤命令；退出条件满足后清旧 Owner。恢复心跳不会恢复旧授权。
    IF NOT xLocked AND xOwnerLost THEN
        nOwner := 0;
        xOwnerLost := FALSE;
        xResetCommands := TRUE;
    END_IF
END_IF

// 同一扫描先处理释放，再按 1/2/3 的优先级处理申请；被拒绝的请求立即应答，不排队自动接管。
FOR i := 1 TO 3 DO
    IF (GVL_control.aStation[i].udiRequestSequence <> 0)
        AND (GVL_control.aStation[i].udiRequestSequence <> GVL_control.aStation[i].udiAckSequence)
        AND (GVL_control.aStation[i].nAction = 2) THEN
        nReply := F_ControlDecision(nOwner := nOwner, nStation := INT_TO_UINT(i), nAction := 2,
            xLocked := xLocked, xOnline := GVL_control.aStation[i].xOnline);
        IF nReply = 1 THEN nOwner := 0; xResetCommands := TRUE; END_IF
        GVL_control.aStation[i].nResult := nReply;
        GVL_control.aStation[i].udiAckSequence := GVL_control.aStation[i].udiRequestSequence;
    END_IF
END_FOR
FOR i := 1 TO 3 DO
    IF (GVL_control.aStation[i].udiRequestSequence <> 0)
        AND (GVL_control.aStation[i].udiRequestSequence <> GVL_control.aStation[i].udiAckSequence) THEN
        nReply := F_ControlDecision(nOwner := nOwner, nStation := INT_TO_UINT(i),
            nAction := GVL_control.aStation[i].nAction, xLocked := xLocked,
            xOnline := GVL_control.aStation[i].xOnline);
        IF (nReply = 1) AND (GVL_control.aStation[i].nAction = 1) THEN
            nOwner := INT_TO_UINT(i);
        END_IF
        GVL_control.aStation[i].nResult := nReply;
        GVL_control.aStation[i].udiAckSequence := GVL_control.aStation[i].udiRequestSequence;
    END_IF
END_FOR
GVL_control.xOwnerChanged := (nOwner <> nOldOwner) OR xResetCommands;
IF GVL_control.xOwnerChanged THEN
    // 清所有站点的旧运动命令，新持有者必须重新下发，不能继承旧按钮或排队动作。
    FOR i := 1 TO 3 DO
        GVL_control.aStation[i].aAxis := aEmpty;
        GVL_control.aStation[i].xWaveSession := FALSE;
    END_FOR
    // 新控制端不得继承上一个站的轨迹触发位。
    GVL_motion.xStart := FALSE;
    GVL_motion.xUpload := FALSE;
    GVL_motion.xAssemble := FALSE;
    GVL_motion.xClear := FALSE;
    GVL_motion.xReset := FALSE;
    GVL_motion.xStop := FALSE;
END_IF
IF nOwner = 0 THEN xOwnerLost := FALSE; END_IF
GVL_control.xCanCommand := FALSE;
FOR i := 1 TO 3 DO
    GVL_control.aStation[i].xGranted := (nOwner = i) AND NOT xOwnerLost AND GVL_control.aStation[i].xOnline;
    GVL_control.xCanCommand := GVL_control.xCanCommand OR GVL_control.aStation[i].xGranted;
END_FOR
GVL_control.nOwner := nOwner;
GVL_control.xLocked := xLocked;
GVL_control.xCanRelease := (nOwner <> 0) AND NOT xLocked AND NOT xOwnerLost;
GVL_control.xStopOwner := xOwnerLost;

END_FUNCTION_BLOCK

// ---- POUs/ControlAuthority_控制权/F_ControlDecision.TcPOU
FUNCTION F_ControlDecision : UINT
// 纯仲裁判定，方便针对真实 ST 条件进行离线边界测试。
VAR_INPUT
    nOwner : UINT; // 当前控制权持有站；0 未分配，1 控制室、2 拖车本地、3 远程室。
    nStation : UINT; // 本次申请或释放的来源站号，合法范围 1～3，站号越小优先级越高。
    nAction : UINT; // 本次控制权操作：1 申请，2 释放。
    xLocked : BOOL; // 统一交接锁；TRUE 时拒绝转交或释放，持有站重复申请仍可确认授权。
    xOnline : BOOL; // 请求来源站心跳在线标志；FALSE 时拒绝该站请求。
END_VAR

// 成功应答不总表示交接：本持有者重复申请只是确认已有权限。
IF (nStation < 1) OR (nStation > 3) OR ((nAction <> 1) AND (nAction <> 2)) THEN
    F_ControlDecision := 7;
ELSIF NOT xOnline THEN
    F_ControlDecision := 4;
ELSIF (nAction = 1) AND (nOwner = nStation) THEN
    F_ControlDecision := 1;
ELSIF xLocked THEN
    // 用户规则：运行中包括高优先级站在内，不能申请接管，也不能主动释放。
    F_ControlDecision := 2;
ELSIF nAction = 2 THEN
    IF nOwner = nStation THEN F_ControlDecision := 1;
    ELSE F_ControlDecision := 5;
    END_IF
ELSIF (nOwner <> 0) AND (nStation > nOwner) THEN
    F_ControlDecision := 6;
ELSE
    F_ControlDecision := 1;
END_IF

END_FUNCTION

// ---- POUs/ManualControl_手动控制/FB_AxisCommandGate.TcPOU
FUNCTION_BLOCK FB_AxisCommandGate
// 每扫描在基础轴块之前调用；只从已授权站点邮箱复制命令，反馈字段不受影响。
VAR_INPUT
    nStation : UINT; // MAIN 已确认的命令来源，0 表示无授权或正在交接。
    nAxis : INT; // MAIN 固定传入与 Data 对应的轴号，范围 1～4。
    xStop : BOOL; // 控制端失联停车请求，独立于普通手动命令许可。
END_VAR
VAR_IN_OUT
    Data : ST_AxisAds; // 对应轴内部命令区；本块只改命令字段，保留反馈字段。
END_VAR
VAR
    Command : ST_AxisCommand; // 仅取本轴邮箱一次，速度和方向从同一份副本提取。
END_VAR

IF (nStation >= 1) AND (nStation <= 3) THEN
    Command := GVL_control.aStation[nStation].aAxis[nAxis];
    Data.xStart := Command.xStart;
    Data.xStop := xStop OR Command.xStop;
    Data.jogz := Command.jogz;
    Data.jogf := Command.jogf;
    Data.gohome := Command.gohome;
    Data.reset := Command.reset;
    Data.lrJogSpeed := Command.lrJogSpeed;
ELSE
    // 无有效站号时不读邮箱，清除上一扫描的请求，同时保留失联停车。
    Data.xStart := FALSE;
    Data.xStop := xStop;
    Data.jogz := FALSE;
    Data.jogf := FALSE;
    Data.gohome := FALSE;
    Data.reset := FALSE;
    Data.lrJogSpeed := 0;
END_IF

END_FUNCTION_BLOCK

// ---- POUs/Trajectory_点位与轨迹/FB_FourAxisTrajectory.TcPOU
FUNCTION_BLOCK FB_FourAxisTrajectory
// 四轴整表轨迹：上位机预检后下发 LREAL 位置点，本块收齐后统一执行。
// 正常流程：0 登记各段 -> 全部下发后 5 统一拼表 -> 0 就绪 -> 10 启动检查 -> 15 首点定位
//           -> 20 开外部给定 -> 30 取点 -> 40 保持末点 -> 60 关闭 -> 70 确认静止 -> 0。
// 异常流程：运动阶段转 50 减速，再经 40/60/70 退出，最后在 90 等待复位。
// 本块每 2 ms 调用一次；使能、点动、回原等基础控制在 FB_AxisControl 中。
// xGroupBusy 占用控制防止两块同时运动，但不能代替设备安全回路。
VAR_INPUT
    xAxesReady : BOOL; // 四轴已使能、回零、静止，供启动和首点定位完成时检查。
    xAbort : BOOL; // 外部联停：许可撤销、撤使能、停止、限位或手动命令冲突。
    nAbortReason : UINT; // MAIN 提供的首个联停原因，0 表示本扫描无联停。
    xAxisFault : BOOL; // 任一轴错误或 NC I/O 反馈无效，拒绝启动或触发联停。
END_VAR
VAR_IN_OUT
    Axes : ARRAY[1..4] OF AXIS_REF; // MAIN 传入的原始轴引用，VAR_IN_OUT 直接操作各 NC 轴接口。
END_VAR
VAR
    // 完整四轴位置表，只由本块分段写入；运行中不再接收上传。
    aPosition : ARRAY[1..4, 0..2099999] OF LREAL; // [轴号, 完整表点号]，所有点号从 0 开始，单位由 NC 配置决定。
    aConfig : ARRAY[1..4] OF ST_AxisConfig; // 启动时锁存参数，首点定位、运行及本次停车使用相同参数。
    aSet : ARRAY[1..4] OF ST_TrajectoryPoint; // 本周期四轴的位置、内部速度和加速度；内部速度用于减速停车。
    aEnable : ARRAY[1..4] OF MC_ExtSetPointGenEnable; // 四个外部给定开启实例；异步执行，等待 NC Enabled 反馈。
    aDisable : ARRAY[1..4] OF MC_ExtSetPointGenDisable; // 四个关闭实例；确认全部退出之前不交回手动。
    aMoveInit : ARRAY[1..4] OF MC_MoveAbsolute; // 四轴各自定位到轨迹首点，全部完成才同步执行位置表。
    aStopInit : ARRAY[1..4] OF MC_Stop; // 外部给定尚未开启时的停车，如取消首点定位。
    rtUpload : R_TRIG; // 本段四轴数据写完后的登记请求上升沿。
    rtAssemble : R_TRIG; // 全部段登记后的独立拼表请求上升沿，不自动启动运动。
    rtClear : R_TRIG; // 清除旧表计数和就绪状态的请求上升沿。
    rtStart : R_TRIG; // 完整位置表就绪后启动轨迹的请求上升沿。
    rtReset : R_TRIG; // 轨迹组故障复位请求上升沿，不复位各 NC 轴故障。
    tmHeartbeat : TON; // 上位机运行心跳超时定时器，启动检查/运动期间 1 秒不变则联停。
    tmEnable : TON; // 四轴外部给定开启阶段超时定时器，限时 5 秒。
    tmMoveInit : TON; // 四轴首点定位阶段超时定时器，限时 60 秒。
    tmExit : TON; // 关闭外部给定及确认退出阶段的超时定时器，限时 5 秒。
    udiLastHeartbeat : UDINT; // 上一扫描上位机运行心跳值，用于检测是否发生变化。
    udiSequence : UDINT; // 当前接收/执行位置表锁存的非零上传序号。
    nCount : UDINT; // 当前整条位置表锁存的单轴总点数，四根轴点数相同。
    nReceived : UDINT; // 已登记的单轴点数，表示段确认进度，不代表已拼入执行表。
    nLoaded : UDINT; // 四轴均已成功拼入执行表的点数。
    nSegment : UDINT; // 当前拼表源段号，从 0 开始，范围 0～20。
    nSegmentPoint : UDINT; // 当前源段内的起始点号，从 0 开始。
    nCopyCount : UDINT; // 本扫描每轴复制点数，受批次、段尾和总表尾三重限制。
    nCopyBytes : UDINT; // 本扫描每轴复制的字节数，等于点数乘 LREAL 大小。
    nSendPoint : UDINT; // 当前轨迹执行取点号，从 0 开始，不是实际到位点号。
    nPrevious : UDINT; // 差分计算前一点索引，首点处夹紧到有效表范围。
    nNext : UDINT; // 差分计算后一点索引，末点处夹紧到有效表范围。
    nHoldCycles : UINT; // 末点静止给定的保持扫描次数，每扫描为 2 ms。
    nStopCycles : UINT; // 减速阶段扫描计数，用于满足该阶段的最少扫描次数。
    nState : UINT; // 轨迹阶段码，数值与上位机监控和故障诊断一致。
    i : INT; // 四轴循环索引，范围 1～4。
    xAllEnabled : BOOL; // 四轴 NC 外部给定均已开启；不是四轴伺服使能汇总。
    xAllDisabled : BOOL; // 四轴外部给定均已关闭，相关开启、关闭和首点停止块均释放 Busy。
    xAllStopped : BOOL; // 四轴 NC 均未处于 Moving 状态；仅为本块此项汇总条件。
    xAllInitDone : BOOL; // 四个首点绝对定位块均输出 Done。
    xMovesIdle : BOOL; // 四个首点定位块均已释放 Busy。
    xEnablePending : BOOL; // 至少一个外部给定开启块仍忙，退出时先等待开启请求结束。
    xFeed : BOOL; // 本扫描需要向四轴发送外部位置给定。
    xValid : BOOL; // 当前轴配置、首点到位或内存复制批次的临时检查结果，每次检查重新赋值。
    xCommandAllowed : BOOL; // 轨迹命令来源为当前有效持有站，且本扫描未发生控制权交接。
    xStopCommand : BOOL; // 当前持有站发出的有效组停止保持命令。
    xUploadRequest : BOOL; // 本扫描获准处理的段登记请求；原始沿已消费后再过滤权限。
    xAssembleRequest : BOOL; // 本扫描获准处理的整表拼接请求。
    xClearRequest : BOOL; // 本扫描获准处理的清表请求。
    xStartRequest : BOOL; // 本扫描获准处理的轨迹启动请求。
    xResetRequest : BOOL; // 本扫描获准处理的轨迹组故障复位请求。
    xNormalStop : BOOL; // 正常人工停止，不作为 1007 故障。
    lrNewVelocity : LREAL; // 当前减速计算的下一扫描速度，单位为 NC 位置单位/秒。
    nBlockAxis : UINT; // 本扫描首个定位/开启块错误的轴，四轴循环结束后统一联停。
    nBlockSource : UINT; // 10=首点定位，11=开启外部给定。
    udiBlockError : UDINT; // 本扫描首个定位/开启块原始错误码，后续轴不能覆盖。
END_VAR
VAR CONSTANT
    // 保留原阶段数值及顺序，供监控和原有区间判断使用。
    cStateIdle : UINT := 0; // 空闲及收段。
    cStateAssemble : UINT := 5; // 拼接已确认的点位段。
    cStateCheckStart : UINT := 10; // 检查轴配置和启动条件。
    cStateMoveToFirstPoint : UINT := 15; // 四轴定位到首点。
    cStateEnableSetpoint : UINT := 20; // 开启外部给定。
    cStateRun : UINT := 30; // 按 2 ms 送点。
    cStateHoldLastPoint : UINT := 40; // 保持末点或停车点。
    cStateDecelerate : UINT := 50; // 减速停车。
    cStateDisableSetpoint : UINT := 60; // 关闭外部给定。
    cStateWaitForStandstill : UINT := 70; // 确认静止并释放组占用。
    cStateFault : UINT := 90; // 等待有效故障复位。
    cDt : LREAL := 0.002; // 单位秒，必须等于 PLC/NC SAF 周期和差分函数周期。
    cMaxPoints : UDINT := 2100000; // 单轴完整表容量，与 aPosition 第二维一致。
    cUploadPoints : UDINT := 100000; // 单轴每段容量，与 GVL_motion.aUpload 第三维一致。
    cCopyPointsPerScan : UDINT := 1024; // 每扫描每轴最多复制 8 KiB；需在目标 PLC 实测任务时间。
END_VAR

// 各 Action 共用本实例变量；运行参数锁存和四轴 MC 实例保持原位。
A01_RequestsAndTimers();
A02_ReadAxisStatus();
A03_ResetAndInterlocks();
// 单一分派：阶段改变后留到下一扫描处理，不能顺序调用三个阶段 Action。
CASE nState OF
cStateIdle, cStateAssemble: A04_ReceiveAndAssemble();
cStateCheckStart, cStateMoveToFirstPoint, cStateEnableSetpoint, cStateRun: A05_PrepareAndRun();
cStateHoldLastPoint, cStateDecelerate, cStateDisableSetpoint, cStateWaitForStandstill: A06_StopAndExit();
END_CASE
// MC 块仍每扫描调用一次，状态发布保持在最后。
A07_CallMotionBlocks();
A08_PublishFeedback();

ACTION A01_RequestsAndTimers:
// 请求、来源站和定时器；写请求沿、诊断首因准备及超时实例。
// 无故障时准备本扫描的诊断位置；故障置位后保持首因，直到有效复位。
IF NOT GVL_motion.xError THEN
    GVL_motion.nFaultAxis := 0;
    GVL_motion.nFaultSource := 0;
    GVL_motion.nFaultState := nState;
    GVL_motion.udiCleanupErrorId := 0;
END_IF
// 1. 上位机操作转为上升沿，防止保持 TRUE 时每扫描重复发起请求。
// 接口顺序：写独立段 -> xUpload 登记 -> 全部段确认 -> xAssemble 统一拼表。
// 原始沿先消费；未授权的保持位不能在以后取得权限时自动变成新请求。
xCommandAllowed := GVL_control.xCanCommand AND NOT GVL_control.xOwnerChanged
    AND (GVL_motion.nCommandStation = GVL_control.nOwner);
xStopCommand := xCommandAllowed AND GVL_motion.xStop;
rtUpload(CLK := GVL_motion.xUpload);
rtAssemble(CLK := GVL_motion.xAssemble);
rtClear(CLK := GVL_motion.xClear);
rtStart(CLK := GVL_motion.xStart);
rtReset(CLK := GVL_motion.xReset);
// Q 是 R_TRIG 的输出，只读取；权限过滤使用独立请求位。
xUploadRequest := rtUpload.Q AND xCommandAllowed;
xAssembleRequest := rtAssemble.Q AND xCommandAllowed;
xClearRequest := rtClear.Q AND xCommandAllowed;
xStartRequest := rtStart.Q AND xCommandAllowed;
xResetRequest := rtReset.Q AND xCommandAllowed;
// 交接或失联使旧表失去启动资格；正在运行时仍走原有联停和退出流程。
IF GVL_control.xOwnerChanged OR NOT GVL_control.xCanCommand THEN
    GVL_motion.xDataReady := FALSE;
    GVL_motion.nUploadStation := 0;
    IF (nState = cStateIdle) OR (nState = cStateAssemble) THEN
        nCount := 0; nReceived := 0; nLoaded := 0; udiSequence := 0; nState := cStateIdle;
    END_IF
END_IF

// 心跳只要变化，TON.IN 就变 FALSE，超时计时复位；连续 1 秒不变则 Q=TRUE。
// 状态 10..40 检查该超时；上传状态 5 不要求心跳，因此可以先上传后开始心跳。
tmHeartbeat(IN := GVL_motion.udiHeartbeat = udiLastHeartbeat, PT := T#1S);
udiLastHeartbeat := GVL_motion.udiHeartbeat;
tmEnable(IN := nState = cStateEnableSetpoint, PT := T#5S);
tmMoveInit(IN := nState = cStateMoveToFirstPoint, PT := T#60S);
tmExit(IN := (nState = cStateDisableSetpoint) OR (nState = cStateWaitForStandstill), PT := T#5S);
IF nState <> cStateDecelerate THEN nStopCycles := 0; END_IF
END_ACTION

ACTION A02_ReadAxisStatus:
// 汇总四轴 NC 状态及 MC 上扫描输出；写六项汇总条件。
// 2. 汇总四轴反馈：AND 从 TRUE 开始，OR 从 FALSE 开始。
// Axis.Status 来自 MAIN 本扫描开头的 ReadStatus。
// 各 MC 块在本块末尾调用，因此这里读到的是它们上一扫描的输出。
xAllEnabled := TRUE;
xAllDisabled := TRUE;
xAllStopped := TRUE;
xAllInitDone := TRUE;
xMovesIdle := TRUE;
xEnablePending := FALSE;
FOR i := 1 TO 4 DO
    xAllEnabled := xAllEnabled AND Axes[i].Status.ExtSetPointGenEnabled;
    // NC 外部给定位为 FALSE 还不够，异步 Enable/Disable 和 Stop.Busy 也要释放。
    // 避免已经交回手动，却仍有上一条异步命令尚未结束。
    xAllDisabled := xAllDisabled AND NOT Axes[i].Status.ExtSetPointGenEnabled
        AND NOT aEnable[i].Busy AND NOT aDisable[i].Busy AND NOT aStopInit[i].Busy;
    xAllStopped := xAllStopped AND NOT Axes[i].Status.Moving;
    xAllInitDone := xAllInitDone AND aMoveInit[i].Done;
    xMovesIdle := xMovesIdle AND NOT aMoveInit[i].Busy;
    xEnablePending := xEnablePending OR aEnable[i].Busy;
END_FOR
END_ACTION

ACTION A03_ResetAndInterlocks:
// 先复位和判断联停，再进入状态机；写首因、停止状态及表资格。
// 复位只清故障；上传完整的位置表保留，新运行仍需使用新的轨迹序号。
// 组复位只清本块故障；各 NC 轴故障仍需通过 Axis1..4.reset 复位。
// 必须已静止、外部给定关闭且相关命令释放，才允许重新进入空闲。
// 未消费序号的上传/启动检查故障可按已确认进度重试；已消费序号需清表并换新序号。
IF xResetRequest AND ((nState = cStateIdle) OR (nState = cStateFault))
    AND xAllStopped AND xAllDisabled AND xMovesIdle THEN
    GVL_motion.xError := FALSE;
    GVL_motion.udiErrorId := 0;
    GVL_motion.nFaultAxis := 0;
    GVL_motion.nFaultSource := 0;
    GVL_motion.nFaultState := 0;
    GVL_motion.udiCleanupErrorId := 0;
    GVL_motion.xDone := FALSE;
    nState := cStateIdle;
END_IF

// 上传阶段不占用轴；启动检查和运动阶段任一轴异常均联停。
// 3. 先判断联停再取点，避免停止条件出现后仍多走一帧。
// 1006=心跳超时，1010=轴错误，1007=停止/联锁/冲突/外部给定意外退出。
// 状态 10 尚未发运动命令，可直接进 90；其他阶段先进 50 减速退出。
// 故障置位后不重复把状态 40 拉回 50，保证末点保持和退出可以完成。
IF (nState >= cStateCheckStart) AND (nState <= cStateHoldLastPoint) AND NOT GVL_motion.xError THEN
    IF xAxisFault OR xAbort OR tmHeartbeat.Q
        OR ((nState >= cStateRun) AND NOT xAllEnabled) THEN
        GVL_motion.xError := TRUE;
        IF tmHeartbeat.Q THEN
            GVL_motion.udiErrorId := 1006;
            GVL_motion.nFaultSource := 7;
        ELSIF xAxisFault THEN
            GVL_motion.udiErrorId := 1010;
            GVL_motion.nFaultSource := 8;
            FOR i := 1 TO 4 DO
                IF Axes[i].Status.Error OR Axes[i].Status.IoDataInvalid
                    OR ((i = 1) AND GVL_axis.Axis1.xError) OR ((i = 2) AND GVL_axis.Axis2.xError)
                    OR ((i = 3) AND GVL_axis.Axis3.xError) OR ((i = 4) AND GVL_axis.Axis4.xError) THEN
                    GVL_motion.nFaultAxis := INT_TO_UINT(i); EXIT;
                END_IF
            END_FOR
        ELSE
            GVL_motion.udiErrorId := 1007;
            IF xAbort THEN GVL_motion.nFaultSource := nAbortReason;
            ELSE GVL_motion.nFaultSource := 9;
            END_IF
        END_IF
        IF nState = cStateCheckStart THEN nState := cStateFault; ELSE nState := cStateDecelerate; END_IF
    END_IF
END_IF

// 人工停止：取消收段/拼表/启动检查，运动阶段从当前给定减速；不人为生成故障。
IF xStopCommand AND NOT GVL_motion.xError THEN
    xNormalStop := TRUE;
    GVL_motion.xDataReady := FALSE;
    GVL_motion.xDone := FALSE;
    IF (nState = cStateIdle) OR (nState = cStateAssemble) OR (nState = cStateCheckStart) THEN
        nCount := 0; nReceived := 0; nLoaded := 0; udiSequence := 0; nState := cStateIdle;
        GVL_motion.xStopped := xAllStopped AND xAllDisabled AND xMovesIdle;
    ELSIF (nState = cStateMoveToFirstPoint) OR (nState = cStateEnableSetpoint) OR (nState = cStateRun) THEN
        nStopCycles := 0;
        nState := cStateDecelerate;
    END_IF
END_IF
END_ACTION

ACTION A04_ReceiveAndAssemble:
// 状态 0/5：收段、清表、拼表和启动请求登记；不推进运动点。
CASE nState OF

cStateIdle: // 空闲：先接收所有独立段，再统一拼表；拼接完成后才允许启动。
    // 清表只清计数和就绪状态，不遍历清零约 134.4 MB 的接收区和执行表。
    // 新轨迹必须从偏移 0 连续覆盖所有有效点，旧数据不会在未收齐时被执行。
    // 同扫描多个请求的优先级为 Clear -> Upload -> Assemble -> Start。
    IF xStopCommand THEN
        // 停止保持期间不接受同扫描上传/拼接/启动请求。
    ELSIF xClearRequest AND xAllDisabled AND xMovesIdle THEN
        xNormalStop := FALSE;
        GVL_motion.xStopped := FALSE;
        GVL_motion.nUploadStation := GVL_control.nOwner;
        nCount := 0;
        nReceived := 0;
        nLoaded := 0;
        udiSequence := 0;
        GVL_motion.xDataReady := FALSE;
        GVL_motion.xDone := FALSE;
    ELSIF xUploadRequest AND NOT GVL_motion.xError THEN
        // 只登记写完的独立段，此处不复制任何位置点。
        // 连续偏移及固定段长共同避免漏段、重复段和错段；先检查范围再做 UDINT 减法。
        IF (GVL_motion.nPointCount < 4) OR (GVL_motion.nPointCount > cMaxPoints)
            OR (GVL_motion.nSampleTimeUs <> 2000) OR (GVL_motion.udiUploadSequence = 0)
            OR (GVL_motion.udiUploadSequence = GVL_motion.udiAcceptedSequence)
            OR (GVL_motion.nUploadCount = 0) OR (GVL_motion.nUploadCount > cUploadPoints)
            OR (GVL_motion.nUploadOffset <> nReceived) THEN
            GVL_motion.udiErrorId := 1001;
            GVL_motion.nFaultSource := 17;
        ELSIF nReceived > GVL_motion.nPointCount THEN
            GVL_motion.udiErrorId := 1001;
            GVL_motion.nFaultSource := 17;
        ELSIF GVL_motion.nUploadCount <> MIN(cUploadPoints, GVL_motion.nPointCount - nReceived) THEN
            GVL_motion.udiErrorId := 1001;
            GVL_motion.nFaultSource := 17;
        ELSIF (nReceived <> 0) AND ((GVL_motion.nPointCount <> nCount)
            OR (GVL_motion.udiUploadSequence <> udiSequence)) THEN
            GVL_motion.udiErrorId := 1001;
            GVL_motion.nFaultSource := 17;
        ELSE
            // 接收确认只表示 PC 已声明本段四轴写完；ADS 数据仍须由 PC 遵守只写一次的约定。
            GVL_motion.nUploadStation := GVL_control.nOwner;
            GVL_motion.xStopped := FALSE;
            xNormalStop := FALSE;
            nCount := GVL_motion.nPointCount;
            udiSequence := GVL_motion.udiUploadSequence;
            nReceived := nReceived + GVL_motion.nUploadCount;
            GVL_motion.xDataReady := FALSE;
        END_IF
        IF GVL_motion.udiErrorId <> 0 THEN
            GVL_motion.xError := TRUE;
            nState := cStateFault;
        END_IF
    ELSIF xAssembleRequest AND NOT GVL_motion.xError THEN
        // 必须收到全部段的确认和独立的完成请求，不能因最后一段到齐就自动拼表或启动。
        IF (nCount < 4) OR (nReceived <> nCount) OR (udiSequence = 0)
            OR (udiSequence = GVL_motion.udiAcceptedSequence)
            OR (GVL_motion.nPointCount <> nCount) OR (GVL_motion.nSampleTimeUs <> 2000)
            OR (GVL_motion.udiUploadSequence <> udiSequence) THEN
            GVL_motion.xError := TRUE;
            GVL_motion.udiErrorId := 1001;
            GVL_motion.nFaultSource := 17;
            nState := cStateFault;
        ELSE
            nLoaded := 0;
            GVL_motion.xDataReady := FALSE;
            GVL_motion.xDone := FALSE;
            nState := cStateAssemble;
        END_IF
    ELSIF xStartRequest AND NOT GVL_motion.xError THEN
        GVL_motion.xDone := FALSE;
        GVL_motion.nCurrentPoint := 0;
        // 点位数值由上位机预检；上传完整只代表表已收齐，不代表轴已到首点。
        // 禁止重放已消费序号，避免旧启动命令重复执行轨迹。
        IF NOT GVL_motion.xDataReady OR (GVL_motion.nUploadStation <> GVL_control.nOwner) OR (nLoaded <> nCount) OR (nCount < 4)
            OR (udiSequence = GVL_motion.udiAcceptedSequence)
            OR (GVL_motion.nPointCount <> nCount) OR (GVL_motion.nSampleTimeUs <> 2000)
            OR (GVL_motion.udiUploadSequence <> udiSequence) THEN
            GVL_motion.udiErrorId := 1001;
            GVL_motion.nFaultSource := 17;
        ELSIF NOT xAxesReady OR NOT xAllDisabled OR NOT xMovesIdle
            OR xAbort OR GVL_motion.xStop OR xAxisFault OR tmHeartbeat.Q THEN
            GVL_motion.udiErrorId := 1004;
            GVL_motion.nFaultSource := 16;
        ELSE
            // 锁存本次运行参数；配置仅应在轴静止且轨迹空闲时修改。
            // 状态 10 仅检查轴配置和就绪，随后进入首点定位。
            aConfig := GVL_motion.aConfig;
            nState := cStateCheckStart;
        END_IF
        IF GVL_motion.udiErrorId <> 0 THEN
            GVL_motion.xError := TRUE;
            nState := cStateFault;
        END_IF
    END_IF

cStateAssemble: // 全部段下发后才进入这里，按段号拼入四轴连续表，PC 不得再改接收区。
    IF (GVL_motion.nPointCount <> nCount) OR (GVL_motion.udiUploadSequence <> udiSequence)
        OR (GVL_motion.nSampleTimeUs <> 2000) OR xUploadRequest OR xClearRequest OR xAssembleRequest THEN
        // 元数据或请求冲突使本次拼接失效；复位后重新 xAssemble，从第 0 点重拼。
        GVL_motion.xError := TRUE;
        GVL_motion.udiErrorId := 1001;
        GVL_motion.nFaultSource := 17;
        nState := cStateFault;
    ELSE
        nSegment := nLoaded / cUploadPoints;
        nSegmentPoint := nLoaded MOD cUploadPoints;
        // 同时限制本拍工作量、剩余总点数和当前段剩余量，短末段也不会越界或串轴。
        nCopyCount := MIN(cCopyPointsPerScan, MIN(nCount - nLoaded, cUploadPoints - nSegmentPoint));
        nCopyBytes := nCopyCount * SIZEOF(aPosition[1, 0]);
        xValid := TRUE;
        FOR i := 1 TO 4 DO
            // 每轴只做一次有界内存复制；源/目标独立，地址每扫描现取，不缓存指针。
            IF MEMCPY(destAddr := ADR(aPosition[i, nLoaded]),
                srcAddr := ADR(GVL_motion.aUpload[nSegment, i, nSegmentPoint]), n := nCopyBytes) <> nCopyBytes THEN
                xValid := FALSE;
            END_IF
        END_FOR
        IF NOT xValid THEN
            GVL_motion.xError := TRUE;
            GVL_motion.udiErrorId := 1012;
            GVL_motion.nFaultSource := 18;
            nState := cStateFault;
        ELSE
            // 四轴本批全部复制成功才推进；最后一批完成后才发布整表就绪。
            nLoaded := nLoaded + nCopyCount;
            IF nLoaded = nCount THEN GVL_motion.xDataReady := TRUE; nState := cStateIdle; END_IF
        END_IF
    END_IF

END_CASE
END_ACTION

ACTION A05_PrepareAndRun:
// 状态 10/15/20/30：检查配置、首点、开启、同步取点；一次只执行当前分支。
CASE nState OF

cStateCheckStart: // 单扫描检查配置与轴就绪；整表数值已由上位机在发送前预检。
    // PLC 不再遍历点位表；保留锁存配置检查，供首点定位、运行及停车使用。
    FOR i := 1 TO 4 DO
        xValid := F_AxisConfigValid(aConfig[i])
            AND (aConfig[i].lrStartTolerance > 0) AND (aConfig[i].lrStartTolerance < 1.0E6)
            AND (aConfig[i].lrInitVelocity > 0) AND (aConfig[i].lrInitVelocity <= aConfig[i].lrMaxVelocity);
        IF NOT xValid THEN
            GVL_motion.udiErrorId := 1002;
            GVL_motion.nFaultAxis := INT_TO_UINT(i);
            GVL_motion.nFaultSource := 15;
            EXIT;
        END_IF
    END_FOR
    IF GVL_motion.udiErrorId <> 0 THEN
        GVL_motion.xError := TRUE;
        nState := cStateFault;
    ELSIF NOT xAxesReady THEN
        GVL_motion.xError := TRUE;
        GVL_motion.udiErrorId := 1004;
        GVL_motion.nFaultSource := 16;
        nState := cStateFault;
    ELSE
        FOR i := 1 TO 4 DO
            aSet[i].lrPosition := aPosition[i, 0];
            aSet[i].lrVelocity := 0;
            aSet[i].lrAcceleration := 0;
        END_FOR
        // 启动检查通过后消费序号；首点定位即使失败，也须换新序号重发。
        GVL_motion.udiAcceptedSequence := udiSequence;
        nSendPoint := 0;
        nState := cStateMoveToFirstPoint;
    END_IF

cStateMoveToFirstPoint: // 参考旧工程 move_init：四轴各自定位到首点，全部完成才激活外部给定。
    // 状态 15 让下方 MoveAbsolute.Execute 产生上升沿，速度用 lrInitVelocity。
    // 四轴定位各自规划，到位时间可不同；全部 Done 并检查实际/设定位置偏差后才同步取点。
    // 超过 60 秒报 1011；停止定位需要 MC_Stop，不能只把 MoveAbsolute.Execute 清零。
    IF tmMoveInit.Q THEN
        GVL_motion.xError := TRUE;
        GVL_motion.udiErrorId := 1011;
        GVL_motion.nFaultSource := 19;
        nState := cStateDecelerate;
    ELSIF xAllInitDone AND xAxesReady THEN
        xValid := TRUE;
        FOR i := 1 TO 4 DO
            IF NOT ((ABS(Axes[i].NcToPlc.ActPos - aPosition[i, 0]) <= aConfig[i].lrStartTolerance)
                AND (ABS(Axes[i].NcToPlc.SetPos - aPosition[i, 0]) <= aConfig[i].lrStartTolerance)) THEN
                IF xValid THEN GVL_motion.nFaultAxis := INT_TO_UINT(i); END_IF
                xValid := FALSE;
            END_IF
        END_FOR
        IF xValid THEN nState := cStateEnableSetpoint;
        ELSE
            GVL_motion.xError := TRUE;
            GVL_motion.udiErrorId := 1004;
            GVL_motion.nFaultSource := 16;
            nState := cStateDecelerate;
        END_IF
    END_IF

cStateEnableSetpoint: // 四轴激活过程中持续送静止首点，共同确认后才推进点号。
    // 状态 20 发起异步外部给定开启请求；等待期间仍送静止首点，不推进点号。
    // 用四根轴的 ExtSetPointGenEnabled 汇总确认，而不是只等其中某个 Enable.Done。
    IF tmEnable.Q THEN
        GVL_motion.xError := TRUE;
        GVL_motion.udiErrorId := 1008;
        GVL_motion.nFaultSource := 20;
        nState := cStateDecelerate;
    ELSIF xAllEnabled THEN nState := cStateRun;
    END_IF

cStateRun: // 位置取点方式与参考工程相同，四轴共用 nSendPoint。
    // 四轴都读取同一个 nSendPoint，每扫描只在四轴循环后推进一次点号。
    // 共享点号保证设定值在同一扫描更新，实际跟随误差由各轴 NC/驱动器反馈决定。
    // 相邻位置点转换为速度/加速度，上位机无需额外下发这两个数组。
    nPrevious := nSendPoint;
    IF nSendPoint > 0 THEN nPrevious := nSendPoint - 1; END_IF
    nNext := MIN(nSendPoint + 1, nCount - 1);
    FOR i := 1 TO 4 DO
        aSet[i] := F_TrajectoryPoint(lrPrevious := aPosition[i, nPrevious],
            lrCurrent := aPosition[i, nSendPoint], lrNext := aPosition[i, nNext],
            xEndpoint := (nSendPoint = 0) OR (nSendPoint = nCount - 1));
    END_FOR
    // 反馈的是本扫描准备送出的点号；递增 nSendPoint 只影响下一次状态 30。
    // 本扫描末尾的 Feed 仍发送已经保存在 aSet 中的当前点。
    GVL_motion.nCurrentPoint := nSendPoint;
    IF nSendPoint = nCount - 1 THEN nHoldCycles := 0; nState := cStateHoldLastPoint;
    ELSE nSendPoint := nSendPoint + 1;
    END_IF

END_CASE
END_ACTION

ACTION A06_StopAndExit:
// 状态 40/50/60/70：保持、减速、关闭和退出；故障 90 等待有效复位。
CASE nState OF

cStateHoldLastPoint: // 末点静止给定保持两个周期，随后关闭外部给定，不强制跳回零位。
    // 正常末点和减速终点都到这里；设定速度已经为 0。
    // 静止点多保持两拍，给 NC 消费最后给定留出时间，再发关闭命令。
    FOR i := 1 TO 4 DO aSet[i].lrAcceleration := 0; END_FOR
    nHoldCycles := nHoldCycles + 1;
    IF nHoldCycles >= 2 THEN nState := cStateDisableSetpoint; END_IF

cStateDecelerate: // 外部轨迹按最后的设定速度减速；首点定位由下方 MC_Stop 停车。
    // 至少经过一次 Stop 调用再退出，覆盖定位请求刚被取消但实际轴仍在运动的情况。
    IF nStopCycles < 2 THEN nStopCycles := nStopCycles + 1; END_IF
    xValid := TRUE;
    FOR i := 1 TO 4 DO
        // 正速度逐步降到 0，负速度逐步升到 0，MAX/MIN 防止跨零反向。
        // 各轴停车减速度独立，停车时刻/距离可能不同，不维持四轴路径比例。
        IF aSet[i].lrVelocity > 0 THEN
            lrNewVelocity := MAX(0, aSet[i].lrVelocity - aConfig[i].lrStopDeceleration * cDt);
        ELSE lrNewVelocity := MIN(0, aSet[i].lrVelocity + aConfig[i].lrStopDeceleration * cDt);
        END_IF
        // 位置用梯形积分：pNew=pOld+(vOld+vNew)/2*dt；加速度=(vNew-vOld)/dt。
        // 从最后给定连续减速，不跳到轨迹末点；本实现未加入 jerk 平滑。
        aSet[i].lrPosition := aSet[i].lrPosition + (aSet[i].lrVelocity + lrNewVelocity) * 0.5 * cDt;
        aSet[i].lrAcceleration := (lrNewVelocity - aSet[i].lrVelocity) / cDt;
        aSet[i].lrVelocity := lrNewVelocity;
        xValid := xValid AND (lrNewVelocity = 0);
    END_FOR
    // 外部给定未退出时 NC 的 Moving 可能仍有效；先结束设定减速，再退出并等待实际静止。
    IF xValid AND xMovesIdle AND (nStopCycles >= 2) THEN nHoldCycles := 0; nState := cStateHoldLastPoint; END_IF

cStateDisableSetpoint: // 等待异步 Enable 结束后再 Disable，防止迟到的 Enable 再次打开轴。
    // xAllDisabled 同时检查 NC 标志和 MC.Busy；关闭失败时保持此状态占用。
    // 复位沿可使下方 Disable 暂时撤请求，下一拍重新产生上升沿进行重试。
    IF xAllDisabled THEN nState := cStateWaitForStandstill; END_IF

// 状态 70：关闭命令完成后，再等实际轴静止及定位命令释放。
// 正常结束才置 xDone；发生过联停/故障则转 90，避免误报正常完成。
// 状态 90 没有 CASE 动作，保留故障，等待上方符合条件的复位沿。
cStateWaitForStandstill:
    IF xAllStopped AND xAllDisabled AND xMovesIdle THEN
        IF GVL_motion.xError THEN nState := cStateFault;
        ELSIF xNormalStop THEN GVL_motion.xStopped := TRUE; nState := cStateIdle;
        ELSE GVL_motion.xDone := TRUE; nState := cStateIdle;
        END_IF
    END_IF

END_CASE
END_ACTION

ACTION A07_CallMotionBlocks:
// 每扫描调用四轴 MC 实例，循环结束统一处理错误；写 MC 输出及清理错误。
// 功能块每周期调用；禁止在四轴循环中途改变公共状态。
// 5. 外部给定实际入口：下面的 Feed、Enable、Disable。
// 状态 20 等开启、30 取点、40 保持、50 减速、60 等关闭，都需要持续更新给定。
// 状态 15 用内部 MoveAbsolute 定位，不执行外部轨迹运动。
// 关闭请求发出后仍送静止点，直到 NC 确认外部给定已关闭。
xFeed := (nState >= cStateEnableSetpoint) AND (nState <= cStateDisableSetpoint);
udiBlockError := 0;
nBlockAxis := 0;
nBlockSource := 0;
FOR i := 1 TO 4 DO
    // A. 首点定位：每轴实例保存自己的 Busy/Done/Error，每扫描都要继续调用。
    // Execute 下降沿不等于立即停止，取消时由下面 MC_Stop 完成停车。
    aMoveInit[i](Axis := Axes[i], Execute := nState = cStateMoveToFirstPoint,
        Position := aPosition[i, 0], Velocity := aConfig[i].lrInitVelocity,
        Acceleration := aConfig[i].lrMaxAcceleration, Deceleration := aConfig[i].lrStopDeceleration);
    // B. 尚未开启外部给定的轴使用 MC_Stop；已开启的轴由状态 50 生成减速给定。
    // 避免外部给定有效时同时用 Stop 和 Feed 争用同一根轴。
    aStopInit[i](Axis := Axes[i], Execute := (nState = cStateDecelerate) AND NOT Axes[i].Status.ExtSetPointGenEnabled,
        Deceleration := aConfig[i].lrStopDeceleration);
    IF xFeed THEN
        // C. 送绝对位置，按确认的调用方式固定速度 0、加速度 2000。
        // Direction 固定为 1，使 NC 在运行、反向和末点保持期间持续采纳位置。
        // PLC 内部仍用 aSet 的速度计算减速停车点位。
        // 该函数返回值不代表本点执行完成，不能用它控制 nSendPoint 递增。
        MC_ExtSetPointGenFeed(Axis := Axes[i],
                            Position := aSet[i].lrPosition,
                            Velocity := 0.0,
                            Acceleration := 2000.0,
                            Direction := 1);
    END_IF
    // D. 开启外部给定：状态 20 的 Execute 上升沿发起异步命令。
    // PositionType=ABSOLUTE；Position 传末点用于目标位置监控，不是让轴立即跑到末点。
    // 轴每拍具体走到哪里，由 Feed.Position 决定；首点定位已由 A 完成。
    // MAX(nCount,1)-1 保证空闲时 nCount=0 也只访问第 0 点，不发生 UDINT 下溢。
                aEnable[i](Axis := Axes[i],
                Execute := nState = cStateEnableSetpoint,
                Position := aPosition[i, MAX(nCount, 1) - 1],
                PositionType := POSITIONTYPE_ABSOLUTE);
    // E. 关闭外部给定：状态 60 请求，先等所有开启请求 Busy 结束。
    // xResetRequest 暂时撤销 Execute，下一拍恢复形成新上升沿，供关闭失败后重试。
    // 确认关闭后还需经过状态 70，才把轴交回基础手动控制。
    aDisable[i](Axis := Axes[i],
                Execute := (nState = cStateDisableSetpoint) AND NOT xEnablePending AND NOT xResetRequest);

    // 四轴仍执行同一阶段；只登记最先出错的轴，循环结束后统一改变状态。
    IF nBlockAxis = 0 THEN
        IF aMoveInit[i].Error AND (nState = cStateMoveToFirstPoint) THEN
            udiBlockError := aMoveInit[i].ErrorID; nBlockAxis := INT_TO_UINT(i); nBlockSource := 10;
        ELSIF aEnable[i].Error AND (nState = cStateEnableSetpoint) THEN
            udiBlockError := aEnable[i].ErrorID; nBlockAxis := INT_TO_UINT(i); nBlockSource := 11;
        END_IF
    END_IF
    // 清理错误单独保存；此前已有故障时不能覆盖原始错误号和来源。
    IF ((aStopInit[i].Error AND (nState = cStateDecelerate)) OR (aDisable[i].Error AND (nState = cStateDisableSetpoint)))
        AND (GVL_motion.udiCleanupErrorId = 0) THEN
        IF nState = cStateDecelerate THEN GVL_motion.udiCleanupErrorId := aStopInit[i].ErrorID;
        ELSE GVL_motion.udiCleanupErrorId := aDisable[i].ErrorID;
        END_IF
        IF GVL_motion.udiCleanupErrorId = 0 THEN GVL_motion.udiCleanupErrorId := 1009; END_IF
        IF NOT GVL_motion.xError THEN
            GVL_motion.udiErrorId := GVL_motion.udiCleanupErrorId;
            GVL_motion.nFaultAxis := INT_TO_UINT(i);
            IF nState = cStateDecelerate THEN GVL_motion.nFaultSource := 12;
            ELSE GVL_motion.nFaultSource := 13;
            END_IF
            GVL_motion.nFaultState := nState;
            GVL_motion.xError := TRUE;
        END_IF
    END_IF
END_FOR
IF nBlockAxis <> 0 THEN
    IF NOT GVL_motion.xError THEN
        GVL_motion.udiErrorId := udiBlockError;
        IF udiBlockError = 0 THEN GVL_motion.udiErrorId := 1010; END_IF
        GVL_motion.nFaultAxis := nBlockAxis;
        GVL_motion.nFaultSource := nBlockSource;
        GVL_motion.nFaultState := nState;
        GVL_motion.xError := TRUE;
    END_IF
    nState := cStateDecelerate;
END_IF
// 退出超时只报错，不强行清 Busy 或改回空闲，防止仍被占用的轴接受新运动。
IF tmExit.Q AND ((nState = cStateDisableSetpoint) OR (nState = cStateWaitForStandstill)) THEN
    IF GVL_motion.udiCleanupErrorId = 0 THEN GVL_motion.udiCleanupErrorId := 1009; END_IF
    IF NOT GVL_motion.xError THEN
        GVL_motion.udiErrorId := 1009;
        GVL_motion.nFaultSource := 14;
        GVL_motion.nFaultState := nState;
        GVL_motion.xError := TRUE;
    END_IF
END_IF
END_ACTION

ACTION A08_PublishFeedback:
// 最后发布接收、拼接、状态和占用反馈；不写运动命令。
// 6. 已接收和已拼接分开发布；只有 xDataReady 才表示完整表可进入启动检查。
GVL_motion.nReceivedCount := nReceived;
GVL_motion.udiReceivedSequence := udiSequence;
GVL_motion.nLoadedCount := nLoaded;
GVL_motion.nState := nState;
GVL_motion.xUploadBusy := nState = cStateAssemble;
GVL_motion.xBusy := (nState >= cStateCheckStart) AND (nState <= cStateWaitForStandstill);
GVL_motion.xRunning := nState = cStateRun;
END_ACTION

END_FUNCTION_BLOCK

// ---- POUs/Trajectory_点位与轨迹/F_TrajectoryPoint.TcPOU
FUNCTION F_TrajectoryPoint : ST_TrajectoryPoint
// 无状态位置差分函数：运行时计算给定，不修改位置表或推进点号。
VAR_INPUT
    lrPrevious : LREAL; // 前一点绝对位置 p[k-1]，单位跟随 NC；边界索引由调用方夹紧。
    lrCurrent : LREAL; // 当前点绝对位置 p[k]，单位跟随 NC，未经角度或丝杆换算。
    lrNext : LREAL; // 后一点绝对位置 p[k+1]，单位跟随 NC。
    xEndpoint : BOOL; // 首点或末点标志，按静止端点处理。
END_VAR
VAR CONSTANT
    cDt : LREAL := 0.002; // 差分采样周期 0.002 秒（2 ms），必须与 PLC/NC SAF 周期一致。
END_VAR

F_TrajectoryPoint.lrPosition := lrCurrent;
// 首尾静止；上位机预检首两点、末两点分别相等。
IF xEndpoint THEN
    F_TrajectoryPoint.lrVelocity := 0;
    F_TrajectoryPoint.lrAcceleration := 0;
ELSE
    // 中心差分：速度=(后点-前点)/(2*dt)，加速度=(后点-2*当前点+前点)/dt²。
    // 位置若用 mm，则导数分别为 mm/s、mm/s²；角度轴同理。
    // 二阶差分会放大位置量化噪声，因此上位机位置表需平滑并通过最大加速度检查。
    F_TrajectoryPoint.lrVelocity := (lrNext - lrPrevious) / (2 * cDt);
    F_TrajectoryPoint.lrAcceleration := (lrNext - 2 * lrCurrent + lrPrevious) / (cDt * cDt);
END_IF

END_FUNCTION

// ---- POUs/Feedback_反馈/FB_HmiFeedback.TcPOU
FUNCTION_BLOCK FB_HmiFeedback
// 在 MAIN 的四个基础轴块之后每扫描调用，只发布状态，不写任何轴命令。
// switch 的机器监控和手动轴反馈使用同一批实际 NC/功能块结果。
VAR
    tmHeartbeat : TON; // PLC 自复位心跳定时器，每约 500 ms 推进一次只读监控心跳。
    udiFault : UDINT; // 本扫描选出的完整故障码；轨迹组优先，其次为第一根故障轴。
    nFaultAxis : UINT; // 故障来源轴号：0 为组故障或无故障，1～4 为对应轴。
    i : INT; // 汇总四轴配置、就绪及故障的循环轴号，范围 1～4。
END_VAR

// 1. 自复位 TON 每约 500 ms 产生一个扫描周期的 Q，不依赖上位机写入。
// 心跳始终更新，不能因待机/故障而停住，否则 switch 会认为反馈已过期。
tmHeartbeat(IN := NOT tmHeartbeat.Q, PT := T#500MS);
IF tmHeartbeat.Q THEN
    IF GVL_HMI.stMonitor.udiHeartbeat = UDINT#4294967295 THEN
        GVL_HMI.stMonitor.udiHeartbeat := 0;
    ELSE
        GVL_HMI.stMonitor.udiHeartbeat := GVL_HMI.stMonitor.udiHeartbeat + 1;
    END_IF
END_IF

// 2. 控制权取仲裁结果，模式按实际状态发布；HMI 只读反馈。
GVL_HMI.stMonitor.nControlOwner := GVL_control.nOwner;
// 模式由实际控制端和轨迹占用决定，不再通过 GVL_pc 中转。
IF GVL_control.nOwner = 0 THEN GVL_HMI.stMonitor.nControlMode := 0;
ELSIF GVL_motion.xBusy THEN GVL_HMI.stMonitor.nControlMode := 2;
ELSE GVL_HMI.stMonitor.nControlMode := 1;
END_IF

// 3. 组故障优先，其次取 Axis1..4 的第一个轴故障。每扫描重算，故障消失就清零。
udiFault := 0;
nFaultAxis := 0;
IF GVL_motion.xError THEN
    udiFault := GVL_motion.udiErrorId;
    nFaultAxis := GVL_motion.nFaultAxis;
ELSIF GVL_axis.Axis1.xError THEN
    udiFault := GVL_axis.Axis1.udiErrorId; nFaultAxis := 1;
ELSIF GVL_axis.Axis2.xError THEN
    udiFault := GVL_axis.Axis2.udiErrorId; nFaultAxis := 2;
ELSIF GVL_axis.Axis3.xError THEN
    udiFault := GVL_axis.Axis3.udiErrorId; nFaultAxis := 3;
ELSIF GVL_axis.Axis4.xError THEN
    udiFault := GVL_axis.Axis4.udiErrorId; nFaultAxis := 4;
END_IF
// 有错误标志但源块尚无错误码时，用 1010 表示轴/控制错误，避免“故障且码为零”。
IF (GVL_motion.xError OR (nFaultAxis <> 0)) AND (udiFault = 0) THEN udiFault := 1010; END_IF
GVL_HMI.udiDetailedFaultCode := udiFault;
GVL_HMI.nFaultAxis := nFaultAxis;
IF udiFault > UDINT#65535 THEN
    GVL_HMI.stMonitor.uiWaveFaultCode := UINT#65535;
ELSE
    GVL_HMI.stMonitor.uiWaveFaultCode := UDINT_TO_UINT(udiFault);
END_IF

// 4. 内部轨迹状态不直接当作页面状态：例如内部 30 对应页面“2 造波中”。
// 停车时先显示“停止中”，实际退出后有故障则显示故障，不把停止请求发送成功当作完成。
IF (GVL_motion.nState = 40) OR (GVL_motion.nState = 50)
    OR (GVL_motion.nState = 60) OR (GVL_motion.nState = 70) THEN
    GVL_HMI.stMonitor.nWaveState := 4;
ELSIF udiFault <> 0 THEN
    GVL_HMI.stMonitor.nWaveState := 7;
ELSIF GVL_motion.nState = 30 THEN
    GVL_HMI.stMonitor.nWaveState := 2;
ELSIF (GVL_motion.nState = 5) OR (GVL_motion.nState = 10)
    OR (GVL_motion.nState = 15) OR (GVL_motion.nState = 20) THEN
    GVL_HMI.stMonitor.nWaveState := 1;
ELSIF GVL_motion.xStopped THEN
    GVL_HMI.stMonitor.nWaveState := 5;
ELSIF GVL_motion.xDone THEN
    GVL_HMI.stMonitor.nWaveState := 6;
ELSE
    GVL_HMI.stMonitor.nWaveState := 0;
END_IF

// 5. 保留原始轨迹诊断；本次只接手动和监控，不新增上位机自动造波写入入口。
GVL_HMI.nTrajectoryState := GVL_motion.nState;
GVL_HMI.nCurrentPoint := GVL_motion.nCurrentPoint;
GVL_HMI.nLoadedCount := GVL_motion.nLoadedCount;
GVL_HMI.nPointCount := GVL_motion.nPointCount;
GVL_HMI.xDataReady := GVL_motion.xDataReady;
GVL_HMI.xTrajectoryBusy := GVL_motion.xBusy;

// 6. 整块接口固定布局，轴反馈从本扫描实际结果集中发布。
// 普通 ADS 读取不声明为跨任务原子快照。
GVL_HMI.stMonitor.nVersion := 4;
GVL_HMI.stMonitor.udiProgramVersion := 2026102401;
GVL_HMI.stMonitor.nBehaviorVersion := 1;
GVL_HMI.stMonitor.nFaultAxis := GVL_motion.nFaultAxis;
GVL_HMI.stMonitor.nFaultSource := GVL_motion.nFaultSource;
GVL_HMI.stMonitor.nFaultState := GVL_motion.nFaultState;
GVL_HMI.stMonitor.udiCleanupErrorId := GVL_motion.udiCleanupErrorId;
GVL_HMI.stMonitor.nByteSize := SIZEOF(GVL_HMI.stMonitor);
GVL_HMI.stMonitor.Axis1.lrActualPosition := GVL_axis.Axis1.lrActualPosition;
GVL_HMI.stMonitor.Axis1.lrSpeed := GVL_axis.Axis1.lrSpeed;
GVL_HMI.stMonitor.Axis1.xHomed := GVL_axis.Axis1.xHomed;
GVL_HMI.stMonitor.Axis1.xError := GVL_axis.Axis1.xError;
GVL_HMI.stMonitor.Axis1.xPositiveLimit := GVL_axis.Axis1.xPositiveLimit;
GVL_HMI.stMonitor.Axis1.xNegativeLimit := GVL_axis.Axis1.xNegativeLimit;
GVL_HMI.stMonitor.Axis1.xOriginSignal := GVL_axis.Axis1.xOriginSignal;
GVL_HMI.stMonitor.Axis1.xEnabled := GVL_axis.Axis1.xEnabled;
GVL_HMI.stMonitor.Axis2.lrActualPosition := GVL_axis.Axis2.lrActualPosition;
GVL_HMI.stMonitor.Axis2.lrSpeed := GVL_axis.Axis2.lrSpeed;
GVL_HMI.stMonitor.Axis2.xHomed := GVL_axis.Axis2.xHomed;
GVL_HMI.stMonitor.Axis2.xError := GVL_axis.Axis2.xError;
GVL_HMI.stMonitor.Axis2.xPositiveLimit := GVL_axis.Axis2.xPositiveLimit;
GVL_HMI.stMonitor.Axis2.xNegativeLimit := GVL_axis.Axis2.xNegativeLimit;
GVL_HMI.stMonitor.Axis2.xOriginSignal := GVL_axis.Axis2.xOriginSignal;
GVL_HMI.stMonitor.Axis2.xEnabled := GVL_axis.Axis2.xEnabled;
GVL_HMI.stMonitor.Axis3.lrActualPosition := GVL_axis.Axis3.lrActualPosition;
GVL_HMI.stMonitor.Axis3.lrSpeed := GVL_axis.Axis3.lrSpeed;
GVL_HMI.stMonitor.Axis3.xHomed := GVL_axis.Axis3.xHomed;
GVL_HMI.stMonitor.Axis3.xError := GVL_axis.Axis3.xError;
GVL_HMI.stMonitor.Axis3.xPositiveLimit := GVL_axis.Axis3.xPositiveLimit;
GVL_HMI.stMonitor.Axis3.xNegativeLimit := GVL_axis.Axis3.xNegativeLimit;
GVL_HMI.stMonitor.Axis3.xOriginSignal := GVL_axis.Axis3.xOriginSignal;
GVL_HMI.stMonitor.Axis3.xEnabled := GVL_axis.Axis3.xEnabled;
GVL_HMI.stMonitor.Axis4.lrActualPosition := GVL_axis.Axis4.lrActualPosition;
GVL_HMI.stMonitor.Axis4.lrSpeed := GVL_axis.Axis4.lrSpeed;
GVL_HMI.stMonitor.Axis4.xHomed := GVL_axis.Axis4.xHomed;
GVL_HMI.stMonitor.Axis4.xError := GVL_axis.Axis4.xError;
GVL_HMI.stMonitor.Axis4.xPositiveLimit := GVL_axis.Axis4.xPositiveLimit;
GVL_HMI.stMonitor.Axis4.xNegativeLimit := GVL_axis.Axis4.xNegativeLimit;
GVL_HMI.stMonitor.Axis4.xOriginSignal := GVL_axis.Axis4.xOriginSignal;
GVL_HMI.stMonitor.Axis4.xEnabled := GVL_axis.Axis4.xEnabled;

// 自动页从同一帧读取确认进度和准备条件，不用写成功冒充就绪。
GVL_HMI.stMonitor.nTrajectoryState := GVL_motion.nState;
GVL_HMI.stMonitor.nReceivedCount := GVL_motion.nReceivedCount;
GVL_HMI.stMonitor.nLoadedCount := GVL_motion.nLoadedCount;
GVL_HMI.stMonitor.nPointCount := GVL_motion.nPointCount;
GVL_HMI.stMonitor.nCurrentPoint := GVL_motion.nCurrentPoint;
GVL_HMI.stMonitor.udiReceivedSequence := GVL_motion.udiReceivedSequence;
GVL_HMI.stMonitor.udiAcceptedSequence := GVL_motion.udiAcceptedSequence;
GVL_HMI.stMonitor.udiErrorId := GVL_motion.udiErrorId;
GVL_HMI.stMonitor.nUploadStation := GVL_motion.nUploadStation;
GVL_HMI.stMonitor.xUploadBusy := GVL_motion.xUploadBusy;
GVL_HMI.stMonitor.xDataReady := GVL_motion.xDataReady;
GVL_HMI.stMonitor.xTrajectoryBusy := GVL_motion.xBusy;
GVL_HMI.stMonitor.xRunning := GVL_motion.xRunning;
GVL_HMI.stMonitor.xDone := GVL_motion.xDone;
GVL_HMI.stMonitor.xError := GVL_motion.xError;
GVL_HMI.stMonitor.xStopped := GVL_motion.xStopped;
GVL_HMI.stMonitor.xAxesStopped := GVL_axis.Axis1.xStopped AND GVL_axis.Axis2.xStopped
    AND GVL_axis.Axis3.xStopped AND GVL_axis.Axis4.xStopped;
GVL_HMI.stMonitor.xMotionPermit := GVL_motion.xMotionPermit;
GVL_HMI.stMonitor.xConfigValid := TRUE;
// 未使能轴的 NC 状态为 Disabled；上传和自动使能前也应允许已停稳的空闲轴。
GVL_HMI.stMonitor.xAxesIdle := GVL_HMI.stMonitor.xAxesStopped
    AND NOT GVL_axis.Axis1.xBusy AND NOT GVL_axis.Axis2.xBusy
    AND NOT GVL_axis.Axis3.xBusy AND NOT GVL_axis.Axis4.xBusy;
GVL_HMI.stMonitor.xAxisFault := GVL_axis.Axis1.xError OR GVL_axis.Axis2.xError
    OR GVL_axis.Axis3.xError OR GVL_axis.Axis4.xError;
// MAIN 已在本扫描应用轴参数，发布时直接从同一个配置来源校验。
FOR i := 1 TO 4 DO
    GVL_HMI.stMonitor.xConfigValid := GVL_HMI.stMonitor.xConfigValid
        AND F_AxisConfigValid(GVL_motion.aConfig[i])
        AND (GVL_motion.aConfig[i].lrInitVelocity > 0)
        AND (GVL_motion.aConfig[i].lrInitVelocity <= GVL_motion.aConfig[i].lrMaxVelocity)
        AND (GVL_motion.aConfig[i].lrStartTolerance >= 0) AND (GVL_motion.aConfig[i].lrStartTolerance < 1.0E12);
    GVL_HMI.stMonitor.xAxesIdle := GVL_HMI.stMonitor.xAxesIdle
        AND (GVL_sy.axis[i].Status.StandStill OR GVL_sy.axis[i].Status.Disabled)
        AND NOT GVL_sy.axis[i].Status.Homing
        AND NOT GVL_sy.axis[i].Status.Stopping AND NOT GVL_sy.axis[i].Status.ExtSetPointGenEnabled
        AND NOT GVL_sy.axis[i].Status.IoDataInvalid;
    GVL_HMI.stMonitor.xAxisFault := GVL_HMI.stMonitor.xAxisFault
        OR GVL_sy.axis[i].Status.Error OR GVL_sy.axis[i].Status.IoDataInvalid;
END_FOR

END_FUNCTION_BLOCK
